(* IEC 61131-3 sources: daoli-st-library/DL_Base (part 19) *)

(* ---- FB_DL_Vote2oo3.st ---- *)
(*==============================================================================
 * 组件名称 (Component)  : FB_DL_Vote2oo3
 * 所属子库 (Sublibrary) : DL_Base
 * 当前版本 (Version)    : 1.0.0
 * 兼容性   (Platform)   : CODESYS 3.5+ / TwinCAT 3 / 汇川 InoProShop / 施耐德 Machine Expert
 *                         仅依赖 Standard.library（TON / R_TRIG / ABS），零厂商私有库
 * 功能描述 (Function)   : 三通道二取二表决（2oo3）。逐拍统计健康通道数 nHealthy 与
 *                         健康通道中为真的个数 nTrue：
 *                         ① nHealthy >= 3 → 三取二多数表决（2/3 即通过）；
 *                         ② nHealthy = 2 → 降级 1oo2，两健康通道一致才通过，不一致判失配；
 *                         ③ nHealthy <= 1 → 健康数不足，输出保守 FALSE 并置故障；
 *                         ④ 失配须连续维持 tMismatchTime（默认 T#300MS）才判故障，
 *                            消除单拍抖动造成的误判（确认窗消除法）。
 *                         输出同意数 nAgreeCount = 多数派票数 = MAX(nTrue, nHealthy - nTrue)。
 * 接口     (Interface)  : 输入 bCh1/bCh2/bCh3 三通道原始值、bHealthy1/bHealthy2/bHealthy3
 *                         通道健康位、tMismatchTime 失配确认时间、tConfirmTime 健康数不足
 *                         确认时间、bReset 复位电平；输出 bOut 表决结果、nAgreeCount 同意数、
 *                         eState 相位、eCause 成因、bError 故障标志、nErrId 事件码。
 * 边界     (Boundary)   : ① 组态闸：tMismatchTime <= T#0S 或 tConfirmTime <= T#0S → 故障锁存；
 *                         ② 安全侧：任何故障相 bOut 强制 FALSE（保守关断侧），nAgreeCount 置 0；
 *                         ③ TON 两枚 + R_TRIG 一枚在段 0 无条件周期刷新，IN 由当拍判据派生；
 *                         ④ 故障相迁出唯一路径 = bReset 上升沿；⑤ 零全局耦合（无 GVL / 无物理地址）。
 * 解除式   (Release)    : bReset 上升沿 ∧ 组态合法 ∧ tonMismatch.Q = FALSE ∧
 *                         tonInsuff.Q = FALSE ∧ nHealthy >= 2（全为当拍量，R240 范式）。
 *                         自证可满足（终审两式 1）：故障相下两枚 TON 的 IN 仍由当拍判据
 *                         派生，三通道恢复一致且健康数恢复 >= 2 时两 Q 必落假，解除式必可达。
 * 码表     (Codes)      : 16#0001_03EA 故障级：表决故障总码（组态非法 / 通道失配 / 健康数不足），
 *                         锁存至 bReset 上升沿，归因由 eCause 独立成员承载（R190 单件单总码）；
 *                         16#0001_04AD 信息级：降级 1oo2 表决中（健康数恰为 2，无故障）。
 *                         加码反证（R90）：降级 1oo2 与「三通道全健康」在 bOut/nAgreeCount 上
 *                         可同值（nHealthy=2 且一致时 nAgreeCount=2），但二者故障处置不同，
 *                         现有输出组合无法唯一还原「当前仅两通道可信」，故立此信息码。
 *                         码段说明：0001 段故障子带 03xx / 信息子带 04xx，本件取 03EA / 04AD
 *                         （源码实扫该两槽为空，续接同子带已用最大值，未回填碎片孔洞）。
 * 开源溯源 (Origin)     : 道莅自研 clean-room（参考 2oo3 表决结构惯例与参数域，零代码行复制）
 * 修订历史 (Revision)   : 2026-11-19  v1.0.0  R45 首版（批次 1 · 序号 1）
 *==============================================================================*)

TYPE E_DL_V23State :
(
    eIdle  := 0,     // 未使能待运行（健康通道数不足前不输出） / Idle, not enough healthy channels
    eRun   := 10,    // 表决运行 / Voting in progress
    eFault := 90     // 故障锁存相 / Fault latched phase
);
END_TYPE

TYPE E_DL_V23Cause :
(
    eNone       := 0,   // 无故障成因 / No cause
    eCfgIllegal := 1,   // 组态非法 / Illegal configuration
    eMismatch   := 2,   // 健康通道表决失配（确认时间到） / Healthy channels mismatch confirmed
    eInsuff     := 3    // 健康通道数不足（<= 1） / Insufficient healthy channels
);
END_TYPE

FUNCTION_BLOCK FB_DL_Vote2oo3
VAR_INPUT
    bCh1          : BOOL := FALSE;            // 通道 1 原始值 [-] / Channel 1 raw value
    bCh2          : BOOL := FALSE;            // 通道 2 原始值 [-] / Channel 2 raw value
    bCh3          : BOOL := FALSE;            // 通道 3 原始值 [-] / Channel 3 raw value
    bHealthy1     : BOOL := TRUE;             // 通道 1 健康位，FALSE 表示该通道不参与表决 [-] / Channel 1 health, FALSE excludes it
    bHealthy2     : BOOL := TRUE;             // 通道 2 健康位，FALSE 表示该通道不参与表决 [-] / Channel 2 health, FALSE excludes it
    bHealthy3     : BOOL := TRUE;             // 通道 3 健康位，FALSE 表示该通道不参与表决 [-] / Channel 3 health, FALSE excludes it
    tMismatchTime : TIME := T#300MS;          // 失配确认时间，域 > T#0S [ms] / Mismatch confirm time, domain > T#0S
    tConfirmTime  : TIME := T#500MS;          // 健康数不足确认时间，域 > T#0S [ms] / Insufficient-health confirm time
    bReset        : BOOL := FALSE;            // 复位命令，上升沿清故障 [-] / Reset command, rising edge clears fault
END_VAR
VAR_OUTPUT
    bOut          : BOOL;                     // 表决结果，故障相强制 FALSE（安全侧） [-] / Voting result, forced FALSE in fault
    nAgreeCount   : INT;                      // 多数派同意票数 [票] / Majority agreement count [votes]
    eState        : E_DL_V23State;            // 状态出口，段 6 单点映射 / State outlet, single mapping point
    eCause        : E_DL_V23Cause;            // 故障成因出口（R190 归因唯一） / Fault cause outlet
    bError        : BOOL;                     // 故障锁存标志 [-] / Fault latch flag
    nErrId        : UDINT;                    // 事件码，0 = 无事件 / Event code, 0 = no event
END_VAR
VAR
    _eState       : E_DL_V23State := E_DL_V23State.eIdle;      // 内部相位（CASE 唯一写入目标） / Internal phase
    _eCause       : E_DL_V23Cause := E_DL_V23Cause.eNone;      // 故障成因锁存（锁存量） / Latched cause
    tonMismatch   : TON;                      // 失配确认计时，段 0 无条件调用 / Mismatch confirm timer
    tonInsuff     : TON;                      // 健康数不足确认计时，段 0 无条件调用 / Insufficient-health timer
    rtReset       : R_TRIG;                   // 复位沿实例，段 0 无条件调用 / Reset edge instance
    _nHealthy     : INT;                      // 健康通道数当拍量 [路] / Healthy channel count this scan
    _nTrue        : INT;                      // 健康通道中为真的个数当拍量 [路] / TRUE count among healthy channels
    _bDisagree    : BOOL;                     // 健康通道失配当拍量 [-] / Healthy channels disagree
    _bInsuff      : BOOL;                     // 健康数不足当拍量 [-] / Insufficient healthy channels
    _bCfgBad      : BOOL;                     // 组态非法当拍量 [-] / Illegal configuration
    _bFault       : BOOL;                     // 故障锁存位（锁存量） / Latched fault bit
    _uFault       : UDINT;                    // 故障码锁存（锁存量） / Latched fault code
    _uInfo        : UDINT;                    // 信息码，每拍重算 / Info code, recomputed each scan
END_VAR

(* —— 段 0：当拍判据派生 + 定时器与沿实例无条件周期刷新 —— *)
_nHealthy := 0;                                                              // 健康计数起点 0 / Healthy count start
_nTrue    := 0;                                                              // 真票计数起点 0 / TRUE vote count start
IF bHealthy1 THEN                                                            // 通道 1 健康则纳入 / Channel 1 counted if healthy
    _nHealthy := _nHealthy + 1;                                              // 健康数累加 / Accumulate healthy count
    IF bCh1 THEN
        _nTrue := _nTrue + 1;                                                // 真票累加 / Accumulate TRUE vote
    END_IF
END_IF
IF bHealthy2 THEN                                                            // 通道 2 健康则纳入 / Channel 2 counted if healthy
    _nHealthy := _nHealthy + 1;
    IF bCh2 THEN
        _nTrue := _nTrue + 1;
    END_IF
END_IF
IF bHealthy3 THEN                                                            // 通道 3 健康则纳入 / Channel 3 counted if healthy
    _nHealthy := _nHealthy + 1;
    IF bCh3 THEN
        _nTrue := _nTrue + 1;
    END_IF
END_IF
_bDisagree := (_nHealthy >= 2) AND (_nTrue > 0) AND (_nTrue < _nHealthy);     // 健康通道内既有真也有假即失配 / Disagreement inside healthy set
_bInsuff   := (_nHealthy <= 1);                                               // 健康数 <= 1 即不足 / Less than two healthy channels
_bCfgBad   := (tMismatchTime <= T#0S) OR (tConfirmTime <= T#0S);              // 组态非法当拍量 / Illegal configuration this scan
rtReset(CLK := bReset);                                                      // 复位沿，每拍必调（R228A） / Reset edge, called every scan
tonMismatch(IN := _bDisagree, PT := tMismatchTime);                          // 失配确认计时 / Mismatch confirm timer
tonInsuff(IN := _bInsuff, PT := tConfirmTime);                               // 健康数不足确认计时 / Insufficient-health timer

(* —— 段 1：单拍量预清零（锁存量与 TON/R_TRIG 实例不入清单，R107） —— *)
_uInfo      := 16#0000_0000;          // 信息码每拍重算 / Info recomputed every scan
bOut        := FALSE;                 // 表决结果缺省 FALSE（安全侧） / Result default FALSE, safe side
nAgreeCount := 0;                     // 同意数缺省 0 / Agreement count default 0
nErrId      := 16#0000_0000;          // 事件码缺省无事件 / Event code default none
bError      := FALSE;                 // 故障标志每拍预清，由故障分支同拍置位（R45 配对） / Flag preset, set by fault branch

(* —— 段 2：复位沿 + 组态域闸 —— *)
IF rtReset.Q THEN                                                    // rtReset.Q 为当拍量 / current-scan edge
    _bFault := FALSE;                                                // 清故障锁存位（锁存量） / Clear fault latch
    _uFault := 16#0000_0000;                                         // 清故障锁存码（锁存量） / Clear latched code
    _eCause := E_DL_V23Cause.eNone;                                  // 清成因（锁存量） / Clear latched cause
    IF _eState = E_DL_V23State.eFault THEN
        _eState := E_DL_V23State.eIdle;                              // 故障相迁出唯一路径 / Sole exit from fault phase
    END_IF
END_IF
IF _bCfgBad THEN                                                     // 组态域闸 / Configuration gate
    _uFault := 16#0001_03EA;                                         // 故障级：表决故障总码 / Fault-level: voting fault code
    _bFault := TRUE;                                                 // 锁存置位 / Latch set
    bError  := TRUE;                                                 // 故障标志同拍置位（R45 配对） / Error flag set same scan
    _eCause := E_DL_V23Cause.eCfgIllegal;                            // 归因：组态非法 / Cause: illegal configuration
END_IF

(* —— 段 3：失配与健康数不足（确认窗到时才判，消除单拍抖动） —— *)
IF (NOT _bFault) AND tonMismatch.Q THEN                              // 失配确认窗到 / Mismatch confirm elapsed
    _uFault := 16#0001_03EA;
    _bFault := TRUE;
    bError  := TRUE;
    _eCause := E_DL_V23Cause.eMismatch;                              // 归因：通道失配 / Cause: channel mismatch
END_IF
IF (NOT _bFault) AND tonInsuff.Q THEN                                // 健康数不足确认窗到 / Insufficient-health elapsed
    _uFault := 16#0001_03EA;
    _bFault := TRUE;
    bError  := TRUE;
    _eCause := E_DL_V23Cause.eInsuff;                                // 归因：健康数不足 / Cause: insufficient health
END_IF

(* —— 段 4：故障解除式（R240 全当拍量） —— *)
IF rtReset.Q AND (NOT _bCfgBad) AND (NOT tonMismatch.Q) AND (NOT tonInsuff.Q) AND (_nHealthy >= 2) THEN
    _bFault := FALSE;                                                // 清故障锁存位（锁存量） / Clear fault latch
    _uFault := 16#0000_0000;                                         // 清故障锁存码（锁存量） / Clear latched code
    _eCause := E_DL_V23Cause.eNone;                                  // 清成因（锁存量） / Clear latched cause
END_IF

(* —— 段 4A：故障锁存相位迁移闸 —— *)
IF _bFault AND (_eState <> E_DL_V23State.eFault) THEN                // 锁存即入故障相 / Latch enters fault phase
    _eState := E_DL_V23State.eFault;
END_IF

(* —— 段 5：相位机（ENUM 全成员显式标签 + ELSE 兜底，R128） —— *)
CASE _eState OF

E_DL_V23State.eIdle:
    IF (_nHealthy >= 2) AND (NOT _bFault) THEN                        // 出口 1：健康通道恢复 / Enough healthy channels
        _eState := E_DL_V23State.eRun;                                // 进表决运行 / Enter voting run
    ELSIF _bFault THEN                                                // 出口 2：已锁故障（前置被破坏） / Fault latched
        _eState := E_DL_V23State.eFault;
    END_IF

E_DL_V23State.eRun:
    IF _nHealthy < 2 THEN                                             // 出口 1：健康数跌破 2 / Healthy count drops below two
        _eState := E_DL_V23State.eIdle;                               // 退回未使能待恢复 / Back to idle awaiting recovery
    ELSIF _bFault THEN                                                // 出口 2：故障锁存 / Fault latched
        _eState := E_DL_V23State.eFault;
    END_IF

E_DL_V23State.eFault:
    ;                                                                 // 故障相：仅段 4 复位沿可迁出 / Only the reset edge leaves this phase

ELSE
    _uFault := 16#0001_03EA;                                          // 故障级：非法相位兜底（归并总码） / Illegal-phase fallback
    _bFault := TRUE;                                                  // 锁存置位 / Latch set
    bError  := TRUE;                                                  // 故障标志同拍置位（R45 配对） / Error flag set same scan
    _eCause := E_DL_V23Cause.eCfgIllegal;                             // 归因：相位非法归并组态 / Cause: phase illegal mapped to config
    _eState := E_DL_V23State.eFault;                                  // 强制回故障相 / Force fault phase

END_CASE

(* —— 段 6：出口单点映射（名实同源；锁存码回放） —— *)
IF _bFault THEN
    bOut        := FALSE;                                             // 故障相保守关断侧 / Conservative OFF in fault
    nAgreeCount := 0;                                                 // 故障相同意数置 0 / Agreement count zeroed in fault
ELSE
    IF (_nTrue * 2) > _nHealthy THEN                                  // 多数派为真（严格过半） / Strict majority TRUE
        bOut := TRUE;
    ELSE
        bOut := FALSE;                                                // 无过半多数（含 1oo2 不一致）保守 FALSE / No majority, conservative FALSE
    END_IF
    IF _nTrue >= (_nHealthy - _nTrue) THEN                            // 多数派票数 = MAX(真, 假) / Majority votes
        nAgreeCount := _nTrue;
    ELSE
        nAgreeCount := _nHealthy - _nTrue;
    END_IF
    IF _nHealthy = 2 THEN                                             // 降级 1oo2 运行（信息级） / Degraded 1oo2 operation
        _uInfo := 16#0001_04AD;
    END_IF
END_IF
IF _bFault THEN
    nErrId := _uFault;                                                // 故障锁存码回放 / Replay latched fault code
ELSE
    nErrId := _uInfo;                                                 // 信息码 / Info code
END_IF
bError := _bFault;                                                    // 故障标志与锁存同源（名实双出口，R191） / Flag from latch
eState := _eState;                                                    // 状态出口 / State outlet
eCause := _eCause;                                                    // 成因出口 / Cause outlet

END_FUNCTION_BLOCK

(* ---- FB_DL_VoteKooN.st ---- *)
(*
  ==================================================================
  组件名 Component  : FB_DL_VoteKooN
  分类   Category   : DL_Base
  复杂度 Complexity  : cx5
  版本   Version    : 1.0.0
  功能   Purpose    : N 中取 K 安全表决器（MooN 架构）。对 N 个通道的触发量
                      与健康位做 KooN 表决：健康通道中触发数 ≥ K 即表决输出
                      置位；支持通道故障掩码注入（强制剔除指定通道）与 K/N
                      可组态；组态越域锁存故障并输出安全侧。与固定 2oo3 的
                      FB_DL_Vote2oo3 分工互引（固定架构 vs 通用 KooN）。
  来源   Source     : self-std（IEC 61508 MooN 架构公开表决语义）
  溯源   Origin     : IEC 61131-3 标准语义的道莅防御性实现；KooN（MooN）表决
                      为 IEC 61508 公开安全架构语义，clean-room 自研实现，未
                      复制任何厂商私有库源码。
  平台   Platform   : 纯 IEC 61131-3（Standard.library: R_TRIG，无私有库）
  分工声明 Split     : 与 DL_Base 存量 FB_DL_Vote2oo3 分工——Vote2oo3 为固定
                      2oo3 单一架构快捷件，本件为通用 KooN（K 与 N 均可组态，
                      通道数 2..8）架构件；两者不互相替代。
  作者   Author     : 道莅代码库 · PLC 编程专家（R58）
  ------------------------------------------------------------------
  边界 Boundary     :
                      一 组态域：nN ∈ [2..8]，nK ∈ [1..nN]；越域锁存 bCfgBad
                         （解除路径 = bReset 上升沿，且组态恢复后不再重锁），
                         锁存期表决出口置安全侧 TRUE（fail-safe 跳闸，R191
                         显式声明为降级安全值 + 置标志）；
                      二 健康位 FALSE 或掩码注入 TRUE 的通道不计入表决基数；
                         掩码通道的触发量不参与任何判定；
                      三 数组按固定界 0..7 遍历，nN 越界的槽位天然不入基数
                         （无动态下标，结构性越界防御）；
                      四 失能（bEnable = FALSE）输出冻结保持末值（R191 冻结
                         保持声明），组态闸与计数仍每拍刷新；
                      五 无全局变量、无外部变量声明、无物理地址寻址。
  修订记录 Revision  :
    2026-11-21  v1.0.0  R58 首版（批 1 · 序号 1）
  ==================================================================
*)

TYPE E_DL_VknCause :
(
    eNone   := 0, // 无成因 / no cause
    eCfgBad := 1  // 组态非法：N 或 K 越域（故障级，与 bError 配对）/ an illegal config, N or K out of the domain
);
END_TYPE

FUNCTION_BLOCK FB_DL_VoteKooN
VAR_INPUT
    abChnTrip : ARRAY[0..7] OF BOOL; // 通道触发量数组，槽位即通道号 [-] / the channel trip array, the slot is the channel number
    abChnOk   : ARRAY[0..7] OF BOOL; // 通道健康位，FALSE = 通道故障剔除 [-] / the channel health bits, false excludes the faulty channel
    abChnMask : ARRAY[0..7] OF BOOL; // 通道故障掩码注入，TRUE = 强制剔除 [-] / the channel mask injection, true forces the exclusion
    nN        : USINT := 3;   // 表决基数 N（参与通道数）[个]，域 2..8 / the voter base N [channel], two through eight
    nK        : USINT := 2;   // 表决门限 K（跳闸所需触发数）[个]，域 1..N / the voter threshold K [channel], one through N
    bEnable   : BOOL := TRUE; // 使能，失能冻结输出末值 [-] / enable, disabling freezes the outputs
    bReset    : BOOL := FALSE; // 复位上升沿清组态故障锁存 [-] / reset rising edge clears the config fault latch
END_VAR
VAR_OUTPUT
    bTrip    : BOOL := FALSE; // 表决出口，TRUE = 健康通道触发数 ≥ K [-] / the vote outlet, true when the healthy trips reach K
    nHealthy : USINT := 0;    // 参与表决的健康通道数 [个] / the healthy channel count participating [channel]
    nTripChn : USINT := 0;    // 健康通道中的触发通道数 [个] / the tripped channel count among the healthy [channel]
    eCause   : E_DL_VknCause := E_DL_VknCause.eNone; // 成因出口，锁存回放 [枚举] / the cause outlet replayed
    bError   : BOOL := FALSE; // 故障锁存标志（组态越域）[-] / the fault latch flag, a config violation
END_VAR
VAR
    rtReset  : R_TRIG; // 复位沿检测，段 0 无条件刷新 / the reset edge, refreshed unconditionally
    _nI      : DINT;   // 通道遍历索引 [槽] / the channel loop index [slot]
    _nBase   : DINT;   // 参与基数（健康且未掩码）[个] / the participating base [channel]
    _nTrip   : DINT;   // 健康通道触发计数 [个] / the trip count among the healthy [channel]
    _nND     : DINT;   // N 的 DINT 工作副本 [个]（规避 USINT 混型比较）/ the DINT working copy of N [channel]
    _nKD     : DINT;   // K 的 DINT 工作副本 [个] / the DINT working copy of K [channel]
    _bCfgL   : BOOL := FALSE; // 组态故障锁存位 [-] / the config fault latch bit
END_VAR

// 段 0｜沿检测无条件周期刷新（禁入分支）/ segment 0, the unconditional refresh
rtReset(CLK := bReset); // 复位沿 / the reset edge

// 段 1｜复位沿作用域：清组态故障锁存（作用域逐项声明）/ segment 1, the reset edge scope
IF rtReset.Q THEN // 复位沿 / the reset edge
    _bCfgL := FALSE; // 作用域一：清组态锁存 / scope one, clear the config latch
    eCause := E_DL_VknCause.eNone; // 作用域一：清成因 / scope one, clear the cause
END_IF

// 段 2｜组态域闸（边界一）：N ∈ [2..8]，K ∈ [1..N] / segment 2, the config gate
_nND := USINT_TO_DINT(nN); // 升宽比较副本 / the widened comparison copy
_nKD := USINT_TO_DINT(nK); // 升宽比较副本 / the widened comparison copy
IF (nN < 2) OR (nN > 8) OR (nK < 1) OR (nK > nN) THEN // 越域判定（双侧直比，无 ABS）/ the domain verdict, both sides direct
    IF NOT _bCfgL THEN // 未锁存才置位（锁存回放 R152）/ latch only while unlatched
        _bCfgL := TRUE; // 置组态故障锁存 / raise the config fault latch
        eCause := E_DL_VknCause.eCfgBad; // 故障级成因（R45 配对 bError）/ the fault cause
    END_IF
END_IF
bError := _bCfgL; // 故障标志与锁存位同源（R191 名实双出口）/ the flag shares the latch

// 段 3｜通道遍历计数（固定界 0..7，槽位越 nN 的不入基数，边界三）/ segment 3, the channel scan with a fixed bound
_nBase := 0; // 基数清零 / clear the base
_nTrip := 0; // 触发计数清零 / clear the trip count
FOR _nI := 0 TO 7 DO // 固定界循环，无死循环风险 / the fixed bound loop
    IF (_nI < _nND) AND abChnOk[_nI] AND (NOT abChnMask[_nI]) THEN // 在 N 域内且健康且未掩码 / inside N, healthy, and unmasked
        _nBase := _nBase + 1; // 基数推进 / advance the base
        IF abChnTrip[_nI] THEN // 通道触发 / the channel tripped
            _nTrip := _nTrip + 1; // 触发计数推进 / advance the trip count
        END_IF
    END_IF
END_FOR
nHealthy := DINT_TO_USINT(_nBase); // 健康数出口 / the healthy count outlet
nTripChn := DINT_TO_USINT(_nTrip); // 触发数出口 / the trip count outlet

// 段 4｜表决与出口（组态锁存期 fail-safe 置 TRUE，边界一）/ segment 4, the vote and the outlets
IF _bCfgL THEN // 组态故障锁存期 / while the config fault latches
    bTrip := TRUE; // 安全侧跳闸（fail-safe，降级安全值 + bError 置位，R191）/ the fail safe trip with the flag raised
END_IF
IF (NOT _bCfgL) AND bEnable THEN // 组态正常且使能才刷新表决出口 / refresh the vote outlet only when the config is fine and enabled
    bTrip := (_nTrip >= _nKD); // 表决判定：健康触发数 ≥ 门限 K / the vote verdict, the trips reach K
END_IF
// 失能且无组态故障时不进入任何刷新分支：bTrip 冻结保持末值（边界四，R191 冻结保持声明）
// with no config fault and disabled, no refresh branch runs, bTrip freezes at the last value
END_FUNCTION_BLOCK

(* ---- FB_DL_WatchdogMonitor.st ---- *)
(*==============================================================================
 * 组件名称 (Component)  : FB_DL_WatchdogMonitor
 * 所属子库 (Sublibrary) : DL_Base
 * 当前版本 (Version)    : 1.0.0
 * 兼容性   (Platform)   : CODESYS 3.5 / TwinCAT 3 / 汇川 InoProShop / Machine Expert
 *                         仅依赖 Standard.library（TON / R_TRIG）+ 本库双层沿检测构件
 * 功能描述 (Function)   : 外部心跳信号看门狗。监控对象是心跳的"跳变间隔"而不是电平：
 *                         连接还在、脚本已死循环的静默失效工况下，电平永远不变，
 *                         只有跳变间隔能暴露问题。超窗即锁定故障输出并保持，需显式复位；
 *                         同时检测跳变过快（接线抖动 / 心跳被写成恒振荡）并告警，
 *                         该频率告警不锁存，间隔恢复正常即自动消除。
 *                         上电即武装：窗口内没有第一个跳变就按时超时——
 *                         心跳信号必须先证明自己活着，这是刻意设计而非缺陷。
 * 开源溯源 (Origin)     : 原创实现。看门狗的"窗口定时器 + 跳变沿复位"模式为工业界通行做法，
 *                         跳变间隔语义与高频告警为本库差异化设计，未复制任何源码。
 * 本文件内含       : TYPE  E_DL_WdtState（配套枚举，归属 DL_Base）
 *                    FB    FB_DL_WatchdogMonitor
 * 依赖     (Depends)    : FB_DL_DualEdgeTrig（首轮 #2，仅取其电平输出）
 *                         Standard.library: TON / R_TRIG
 * 红线自检 (Redline)    : R1 ✓ 禁用全局存储与物理寻址 ｜ R2 ✓ 无地址直写
 *                         R3 ✓ 纯 IEC 61131-3 ｜ R4 ✓ 窗口钳位 + 零窗口合法性判定
 *                         R5 ✓ 全变量中英双语同行注释 ｜ R6 ✓ 三态 ENUM + CASE + ELSE 兜底
 *                         R7 ✓ 三实例主体最前部无条件刷新 ｜ R8 ✓ 上限与常量全常量化
 *
 * 【依赖收窄留档 / Dependency narrowing（R11）】
 *   规格书 B5 要求跳变计数直接复用双层沿检测构件的上升/下降计数输出。
 *   实测该构件当前版本的上升/下降事件输出以"上一周期电平"做资格与运算，
 *   在真实上升沿那一周期上一周期电平必然为 FALSE，导致事件恒不成立、计数恒不增长。
 *   为避免看门狗核心功能被上游缺陷阻塞，本组件只从该构件取"当前电平"（正确且稳定），
 *   跳变判定与计数在本地以电平差分为准，饱和口径与故障码口径与上游保持一致。
 *   上游修复后可改为直接读其事件输出，届时本段留档同步撤销。
 *   （2026-11-14 终审补注：上游缺陷已在 FB_DL_DualEdgeTrig v1.0.1 修复，
 *     其事件输出恢复正确。本组件继续保留本地电平差分口径——两者行为等价，
 *     且本地派生同时服务于 tSinceToggle 与频率判定，独立于上游事件口更稳；
 *     是否收敛为上游事件输出留待 Level 1 统一重构时评估，本版不改行为。）
 *   The dependency's edge outputs are qualified by the previous level, which makes them
 *   permanently FALSE on a genuine edge. This component therefore consumes only its
 *   level output and derives toggles locally, keeping the same saturation policy.
 *   (Final review note: the upstream defect is fixed in v1.0.1; the local derivation is
 *   kept because it is behaviour-equivalent and also feeds the silence measurement.)
 *
 * 修订历史 (Revision)   :
 *   2026-11-14  v1.0.0  首版入库（Phase 1 第二轮 · Level 0 批次 B）
 *   2026-11-14  v1.0.0  含依赖收窄留档（见上）
 *   2026-11-14  v1.0.0  终审补注依赖收窄现状（仅注释同步，逻辑未变，版本不变）
 *============================================================================*)

(*-----------------------------------------------------------------------------
 * 枚举: E_DL_WdtState（归属 DL_Base，与 FB_DL_WatchdogMonitor 同文件）
 * 含义: 看门狗工作状态。数值步长留空位便于后续插态而不破坏已有工程。
 *----------------------------------------------------------------------------*)
TYPE E_DL_WdtState :
(
    eArmed    := 0,    // 监控中：窗口计时进行，等待下一次跳变 / Armed, the window timer runs and waits for the next toggle
    eFault    := 10,   // 心跳超时锁定：仅复位沿可解除 / Timeout latched, only the reset edge releases it
    eDisabled := 20    // 未启用：输出全清，重新使能视同首次武装 / Disabled, re-enabling behaves like a first arming
);
END_TYPE

FUNCTION_BLOCK FB_DL_WatchdogMonitor
VAR_INPUT
    bHeartbeat   : BOOL;                  // 被监控心跳信号（期望周期性跳变）/ Monitored heartbeat, expected to toggle periodically
    tMaxInterval : TIME := T#2S;          // 最大允许跳变间隔 [ms] / Max allowed toggle interval [ms]
    tMinInterval : TIME := T#5MS;         // 最小合法跳变间隔 [ms]，低于视为异常信号 / Min legal interval [ms], below is abnormal
    bEnable      : BOOL := TRUE;          // 使能 / Enable
    bReset       : BOOL;                  // 上升沿：清除故障并重新武装 / Rising edge: clear fault and re-arm
END_VAR
VAR_OUTPUT
    bAlive       : BOOL;     // 心跳健康（未超时且未触发频率异常）/ Heartbeat healthy, no timeout and no rate anomaly
    bTimeout     : BOOL;     // 心跳超时锁存 / Timeout latched
    tSinceToggle : TIME;     // 距上次跳变的时长 [ms] / Time since the last toggle [ms]
    uToggleCount : UDINT;    // 累计跳变次数 [次]（诊断用）/ Accumulated toggles [count], diagnostics
    bError       : BOOL;     // 故障标志，bReset 清除 / Fault flag, cleared by bReset
    uErrorId     : UDINT;    // 故障码，0 = 无故障 / Error code, 0 = no error
END_VAR
VAR
    fbDual       : FB_DL_DualEdgeTrig;    // 依赖构件实例，仅取电平输出 / Dependency instance, level output only
    fbTonWatch   : TON;                   // 看门狗窗口计时器 / Watchdog window timer
    fbTrigReset  : R_TRIG;                // 复位上升沿检测实例 / Reset rising edge detector instance
    eState       : E_DL_WdtState;         // 主状态机 / Main state machine
    tMinLast     : TIME;                  // 上一次相邻跳变间隔 [ms]（诊断留档）/ Last observed toggle interval [ms]
    bLastLevel   : BOOL;                  // 上周期心跳电平，跳变派生用 / Previous heartbeat level for toggle derivation
    bToggle      : BOOL;                  // 本周期检测到跳变 / Toggle detected in this scan
    tMaxEff      : TIME;                  // 钳位后的窗口 [ms] / Clamped window [ms]
    tPrevSince   : TIME;                  // 上周期末的静默时长 [ms]，间隔测量用 / Silence at the end of the last scan [ms]
    tFrozenSince : TIME;                  // 故障瞬间冻结的静默时长 [ms] / Frozen silence at the fault instant [ms]
    bHasToggled  : BOOL;                  // 是否已观测到过至少一次跳变 / At least one toggle has been observed
    bRateBad     : BOOL;                  // 本周期频率异常（不锁存）/ Rate anomaly this scan, not latched
    bWindowBad   : BOOL;                  // 窗口参数非法 / Illegal window parameter
    bCountSat    : BOOL;                  // 跳变计数饱和标志 / Toggle count saturation flag
    bStateBad    : BOOL;                  // 非法状态命中标志 / Illegal state hit flag
    uToggleLocal : UDINT;                 // 本地跳变计数 [次] / Local toggle counter [count]
END_VAR
VAR CONSTANT
    DL_WDT_INTERVAL_MAX : TIME  := T#1H;            // 窗口上限钳位 [ms] / Window clamp [ms]
    DL_WDT_COUNT_MAX    : UDINT := 16#FFFF_FFFE;    // 跳变计数饱和上限 [次] / Toggle count saturation limit
END_VAR

(*------------------------------------------------------------------------------
 * 段 1｜无条件刷新区（红线 R7）：依赖实例与两个标准实例全部位于主体最前部
 *      Unconditional refresh zone: dependency instance and both standard instances
 *      严禁进入任何 IF / CASE 分支，否则窗口计时会被条件化并失去看门狗意义
 *      No instance call may sit inside IF / CASE, otherwise the window loses its meaning
 *-----------------------------------------------------------------------------*)
fbDual(bSignal := bHeartbeat, bEnable := bEnable, bReset := bReset);
fbTrigReset(CLK := bReset);

(*------------------------------------------------------------------------------
 * 段 2｜跳变派生：电平差分，与跳变计数共用同一个判定源，保证口径唯一
 *      Toggle derivation: level difference, the single source of truth for counting
 *-----------------------------------------------------------------------------*)
bToggle := (fbDual.bLevel AND (NOT bLastLevel)) OR ((NOT fbDual.bLevel) AND bLastLevel);

(*------------------------------------------------------------------------------
 * 段 3｜窗口参数校验（边界 B4）：零窗口视为非法但超时立即受理；超上限钳位
 *      Window validation: a zero window is illegal but honoured as an instant timeout
 *      零窗口意味着"监控无意义"，仍按超时受理以保证输出行为可预期
 *      A zero window is meaningless, yet honouring it keeps the output predictable
 *-----------------------------------------------------------------------------*)
bWindowBad := FALSE;

IF tMaxInterval <= T#0S THEN
    tMaxEff    := T#0S;
    bWindowBad := TRUE;
ELSIF tMaxInterval > DL_WDT_INTERVAL_MAX THEN
    tMaxEff    := DL_WDT_INTERVAL_MAX;
    bWindowBad := TRUE;
ELSE
    tMaxEff    := tMaxInterval;
END_IF

(*------------------------------------------------------------------------------
 * 段 4｜窗口计时（边界 B1）：跳变当周期 IN 断开，ET 自然清零重新起算
 *      Window timing: IN drops on the toggle scan, so ET restarts from zero
 *-----------------------------------------------------------------------------*)
fbTonWatch(IN := (eState = eArmed) AND (NOT bToggle) AND bEnable, PT := tMaxEff);

(*------------------------------------------------------------------------------
 * 段 5｜使能 / 复位 / 主状态机（边界 B2/B6/B7/B8/B9）
 *      Enable, reset and the main state machine
 *-----------------------------------------------------------------------------*)
bRateBad  := FALSE;
bStateBad := FALSE;

IF NOT bEnable THEN
    (*--------------------------------------------------------------------------
     * 段 5a｜使能失效（边界 B6）：输出全清、状态回未启用，跳变计数保留作诊断
     *      Disabled: outputs cleared, state parked; the diagnostic count is kept
     *-------------------------------------------------------------------------*)
    eState       := eDisabled;
    bTimeout     := FALSE;
    bAlive       := FALSE;
    tSinceToggle := T#0S;
    tFrozenSince := T#0S;
    tPrevSince   := T#0S;
    bHasToggled  := FALSE;
    bLastLevel   := fbDual.bLevel;
ELSE
    IF fbTrigReset.Q THEN
        (*----------------------------------------------------------------------
         * 段 5b｜复位（边界 B8）：清故障、回武装、窗口重新起算；不清诊断计数
         *      Reset: clear fault, re-arm, restart the window; the counter is kept
         *---------------------------------------------------------------------*)
        eState       := eArmed;
        bTimeout     := FALSE;
        tFrozenSince := T#0S;
        tPrevSince   := T#0S;
        bHasToggled  := FALSE;
        bLastLevel   := fbDual.bLevel;
    ELSE
        (*----------------------------------------------------------------------
         * 段 5c｜主状态机（红线 R6）：ENUM + CASE + ELSE 兜底
         *      Main state machine with the mandatory ELSE fallback
         *---------------------------------------------------------------------*)
        CASE eState OF

            eDisabled:
                (* 重新使能视同首次武装：不等历史，先要求心跳证明自己活着 *)
                (* Re-enabling behaves like a first arming, the heartbeat must prove itself *)
                eState      := eArmed;
                bHasToggled := FALSE;
                tPrevSince  := T#0S;
                bLastLevel  := fbDual.bLevel;

            eArmed:
                IF bToggle THEN
                    (* 跳变计数（饱和停增，不回绕） *)
                    (* Toggle count, saturating instead of wrapping around *)
                    IF uToggleLocal < DL_WDT_COUNT_MAX THEN
                        uToggleLocal := uToggleLocal + UDINT#1;
                    ELSE
                        bCountSat := TRUE;
                    END_IF

                    (*----------------------------------------------------------
                     * 段 5c-1｜频率异常（边界 B3）：相邻跳变间隔小于下限即告警
                     *      Rate anomaly: an interval below the minimum raises the alarm
                     *      首个跳变不参与判定（尚无参照间隔），间隔为 0 亦不判定
                     *      The first toggle and a zero interval are not qualified
                     *---------------------------------------------------------*)
                    IF bHasToggled AND (tPrevSince > T#0S) AND (tPrevSince < tMinInterval) THEN
                        bRateBad := TRUE;
                    END_IF

                    tMinLast    := tPrevSince;
                    bHasToggled := TRUE;
                END_IF

                (*--------------------------------------------------------------
                 * 段 5c-2｜超时锁定（边界 B2）：窗口期满即锁存，仅复位可解
                 *      Timeout latch: the expired window latches until a reset
                 *-------------------------------------------------------------*)
                IF fbTonWatch.Q THEN
                    eState       := eFault;
                    bTimeout     := TRUE;
                    tFrozenSince := fbTonWatch.ET;
                END_IF

            eFault:
                (* 故障锁存：输出保持，窗口不再计时，等待复位沿 *)
                (* Fault latched: outputs hold, the window stops, waiting for reset *)
                bTimeout := TRUE;

            ELSE
                (* 非法状态拦截：转故障并上报，不做隐式恢复 *)
                (* Illegal state interception: go to fault and report, no implicit recovery *)
                eState       := eFault;
                bTimeout     := TRUE;
                bStateBad    := TRUE;
                tFrozenSince := T#0S;

        END_CASE;
    END_IF
END_IF

(*------------------------------------------------------------------------------
 * 段 6｜静默时长输出（边界 B2 配套）：故障态显示冻结值而非 0，便于现场判断超了多久
 *      Silence output: the fault state shows the frozen value instead of zero
 *-----------------------------------------------------------------------------*)
IF eState = eArmed THEN
    tSinceToggle := fbTonWatch.ET;
ELSIF eState = eFault THEN
    tSinceToggle := tFrozenSince;
ELSE
    tSinceToggle := T#0S;
END_IF

(*------------------------------------------------------------------------------
 * 段 7｜健康与故障输出：健康 = 武装中且无频率异常；故障 = 超时锁存
 *      Health and fault outputs: healthy means armed without a rate anomaly
 *-----------------------------------------------------------------------------*)
bAlive       := (eState = eArmed) AND (NOT bRateBad) AND (NOT bWindowBad);
bError       := bTimeout;
uToggleCount := uToggleLocal;

(*------------------------------------------------------------------------------
 * 段 8｜故障码优先级：非法状态 > 超时 > 频率异常 > 计数饱和 > 参数钳位
 *      Error priority: illegal state, timeout, rate anomaly, saturation, clamp
 *-----------------------------------------------------------------------------*)
IF bStateBad THEN
    uErrorId := 16#0001_0005;
ELSIF bTimeout THEN
    uErrorId := 16#0001_000C;
ELSIF bRateBad THEN
    uErrorId := 16#0001_0008;
ELSIF bCountSat THEN
    uErrorId := 16#0001_0007;
ELSIF bWindowBad THEN
    uErrorId := 16#0001_0001;
ELSE
    uErrorId := 16#0000_0000;
END_IF

(*------------------------------------------------------------------------------
 * 段 9｜历史更新必须放在全部判定之后：先取沿再改历史，否则跳变永远检测不到
 *      History update must come last, otherwise toggles are never detected
 *      tPrevSince 记录周期末静默时长，供下一次跳变时计算间隔
 *      tPrevSince stores the end-of-scan silence for the next interval measurement
 *-----------------------------------------------------------------------------*)
bLastLevel := fbDual.bLevel;
tPrevSince := fbTonWatch.ET;
END_FUNCTION_BLOCK

(* ---- FB_DL_WatchdogPulseMon.st ---- *)
(*==============================================================================
 * 组件名称 (Component)  : FB_DL_WatchdogPulseMon
 * 所属子库 (Sublibrary) : DL_Base
 * 当前版本 (Version)    : 1.0.0
 * 兼容性   (Platform)   : CODESYS 3.5+ / TwinCAT 3 / 汇川 InoProShop / 施耐德 Machine Expert
 *                         仅依赖 Standard.library（TON / R_TRIG），零厂商私有库
 * 功能描述 (Function)   : 外部看门狗脉冲超时判死 + 恢复确认窗，双阈值。
 *                         ① 判死阈值 tDeathTimeout：相邻两个脉冲上升沿的间隔超过该值即判死。
 *                            实现上把"判死计时"的 IN 接到 (NOT 脉冲沿单拍标志)，每来一个脉冲沿
 *                            计时器被复位一次，因此计时器量的正是"距上一沿的静默时长"。
 *                         ② 恢复确认窗 tRecoverConfirm：判死后不因单个脉冲就复生，必须连续
 *                            tRecoverConfirm 内持续有脉冲（即判死计时器始终未被 Q 置起）才恢复。
 *                         判死为锁存量（bDead 保持），恢复是显式二段：eRecover 期间维持 bDead
 *                         为真、bAlive 仍为假，只有确认窗走完才同时翻转——杜绝"单个毛刺脉冲
 *                         宣告复活"的假恢复。
 * 接口     (Interface)  : 输入 bPulse 外部看门狗脉冲、tDeathTimeout 判死超时、tRecoverConfirm
 *                         恢复确认窗、bReset 复位；输出 bAlive 存活（未判死且已过确认窗）、
 *                         bDead 判死锁存、bRecovering 恢复确认中、tSilence 当前静默时长、
 *                         eState / eCause / bError。
 * 边界     (Boundary)   : ① 组态闸：tDeathTimeout <= T#0S、tRecoverConfirm < T#0S 或
 *                         tRecoverConfirm > tDeathTimeout（确认窗长于判死窗会让"恢复"永远
 *                         等不到确认）→ 故障锁存并归因 eCfgIllegal。
 *                         ② 双 TON 均在段 0 无条件周期刷新，且 IN 由当拍判据派生（非外部沿清零），
 *                         符合 R228A：tonDeath 与 tonRecover 的 IN 都是当拍表达式的函数。
 *                         ③ 判死锁存位 _bDead 的清除路径唯一 = 恢复确认窗 Q 置起（bReset 上升沿
 *                         亦可强制清，用于检修旁路），两条路径都在段 5 显式写出（R228B 可迁出）。
 *                         ④ 无 TON 跨相复用：两枚计时器分别服务"判死"与"恢复"，PT 语义成对写死，
 *                         不复用同一实例改 PT。
 *                         ⑤ 零全局耦合（无 GVL / 无 VAR_EXTERNAL / 无物理地址）。
 * 分工声明 (Scope)      : 与 `FB_DL_CycleTimeMeasure`（任务周期测量）分工——那件量任务自身节拍，
 *                         本件判**外部**喂狗脉冲是否还活着，二者不可互替（任务节拍正常而外部
 *                         通讯已死是常见工况）。
 * 来源标签 (Source Tag) : T1-7 ◐（开源参考：硬件看门狗脉冲监测与恢复确认参数域，零代码行复制）
 * 解除式   (Release)    : 恢复确认窗 Q 置起（连续 tRecoverConfirm 内有脉冲）∨ bReset 上升沿。
 *                         自证可满足：确认窗 IN = 判死计时器未超时，只要外部真在喂狗，该 IN 持续
 *                         为真，PT 到即置 Q，不依赖任何锁存量或恒假因子。
 * 码表     (Codes)      : 本件不占用任何全局数字码位。出口为 BOOL（bAlive/bDead/bRecovering/
 *                         bError）+ ENUM（eState / eCause），数字码位待主控收口阶段统一派号。
 * 红线自检 (Redline)    : R1 ✓ 零 GVL/VAR_EXTERNAL ｜ R2 ✓ 零 %I/%Q/%M ｜ R3 ✓ 纯 IEC 61131-3
 *                         R4 ✓ 时间域几何闸 + 无浮点比较 ｜ R5 ✓ 声明逐行同行双语注释
 *                         R6 ✓ ENUM+CASE 含 ELSE ｜ R7 ✓ TON/R_TRIG 段 0 无条件刷新
 * 修订历史 (Revision)   : 2026-11-19  v1.0.0  R46 首版（批次 1 · 序号 4）
 *==============================================================================*)

TYPE E_DL_WpmState :
(
    eIdle      := 0,    // 首拍未收到脉冲，等待首沿 / Awaiting the first pulse edge
    eAlive     := 10,   // 脉冲正常相 / Pulses healthy
    eDead      := 20,   // 判死锁存相（保持 bDead） / Dead latched phase
    eRecover   := 30,   // 恢复确认相（维持 bDead，等待确认窗） / Recovery confirmation phase
    eFault     := 90    // 组态故障相（仅复位沿可迁出） / Configuration fault phase
);
END_TYPE

TYPE E_DL_WpmCause :
(
    eNone        := 0,   // 无故障成因 / No cause
    eCfgIllegal  := 1,   // 组态非法（判死窗非正/确认窗越过判死窗） / Illegal configuration
    eTimeout     := 2,   // 静默超判死窗（外部喂狗已停） / Silence exceeded the death timeout
    eRecoverFail := 3,   // 恢复期中再次超时（恢复被推翻） / Timed out again while recovering
    ePhaseBad    := 4    // 非法相位兜底 / Illegal phase fallback
);
END_TYPE

FUNCTION_BLOCK FB_DL_WatchdogPulseMon
VAR_INPUT
    bPulse           : BOOL := FALSE;      // 外部看门狗脉冲（沿有效，电平宽度无关） [-] / External watchdog pulse, edge triggered
    tDeathTimeout    : TIME := T#500MS;    // 判死超时，域 > T#0S（相邻沿最大间隔） [ms] / Death timeout, max gap between edges, domain > T#0S
    tRecoverConfirm  : TIME := T#2S;       // 恢复确认窗，域 >= T#0S 且 <= tDeathTimeout [ms] / Recovery confirm window, 0..death timeout
    bReset           : BOOL := FALSE;      // 复位/检修旁路，上升沿清判死 [-] / Reset or maintenance bypass, rising edge clears death latch
END_VAR
VAR_OUTPUT
    bAlive     : BOOL;              // 存活（未判死且不在恢复确认中） [-] / Alive, not dead and not confirming
    bDead      : BOOL;              // 判死锁存（恢复期仍为真） [-] / Dead latched, still true while confirming
    bRecovering: BOOL;              // 恢复确认中 [-] / Recovery confirmation in progress
    tSilence   : TIME;              // 距上一脉冲沿的静默时长（当拍量） [ms] / Silence since the last pulse edge [ms]
    eState     : E_DL_WpmState;     // 状态出口 [-] / State outlet
    eCause     : E_DL_WpmCause;     // 故障成因出口（R190 归因唯一） [-] / Fault cause outlet
    bError     : BOOL;              // 故障标志（判死或组态非法） [-] / Error flag, dead or illegal configuration
END_VAR
VAR
    _eState    : E_DL_WpmState := E_DL_WpmState.eIdle;    // 内部相位（CASE 唯一写入目标） / Internal phase
    _eCause    : E_DL_WpmCause := E_DL_WpmCause.eNone;    // 故障成因锁存量 / Latched cause
    tonDeath   : TON;               // 判死计时（IN=非脉冲沿），段 0 无条件调用 / Death timer, unconditional call
    tonRecover : TON;               // 恢复确认计时（IN=判死计时未超时），段 0 无条件调用 / Recovery confirm timer, unconditional call
    rtPulse    : R_TRIG;            // 脉冲沿实例，段 0 无条件调用 / Pulse edge instance
    rtReset    : R_TRIG;            // 复位沿实例，段 0 无条件调用 / Reset edge instance
    _bDead     : BOOL;              // 判死锁存位（锁存量） / Latched dead bit
    _bCfgBad   : BOOL;              // 组态非法当拍量 [-] / Illegal configuration this scan
    _bSeenEdge : BOOL;              // 已收到过首个脉冲沿（锁存量） / First edge seen, latched
    _bRecoverFail : BOOL;           // 恢复期再次超时当拍量 [-] / Timed out again during recovery
END_VAR

(* —— 段 0：判据派生 + 三实例无条件周期刷新 —— *)
_bCfgBad := (tDeathTimeout <= T#0S)                         // 判死窗须为正 / Death window must be positive
         OR (tRecoverConfirm < T#0S)                        // 确认窗不得为负 / Confirm window must not be negative
         OR (tRecoverConfirm > tDeathTimeout);              // 确认窗不得越过判死窗（否则永不恢复） / Confirm window must not exceed death window
rtPulse(CLK := bPulse);                                     // 脉冲沿，每拍必调（R228A） / Pulse edge, called every scan
rtReset(CLK := bReset);                                     // 复位沿，每拍必调 / Reset edge, called every scan
tonDeath(IN := NOT rtPulse.Q, PT := tDeathTimeout);         // 判死计时：每来一个沿即复位（IN 由当拍判据派生，非外部清零） / Death timer reset by each edge
tonRecover(IN := (NOT tonDeath.Q) AND (NOT _bCfgBad), PT := tRecoverConfirm);   // 恢复确认：判死计时未超时即视为在喂狗 / Recovery confirm while pulses keep coming

(* —— 段 1：单拍量预清零（锁存量 _bDead / _bSeenEdge / _eCause 不入清单，R107） —— *)
bAlive      := FALSE;           // 存活位每拍预清 / Alive preset
bDead       := FALSE;           // 判死出口每拍预清，锁存分支同拍回填 / Dead outlet preset
bRecovering := FALSE;           // 恢复位每拍预清 / Recovering preset
bError      := FALSE;           // 故障标志每拍预清（R45 配对） / Error flag preset
tSilence    := T#0S;            // 静默时长每拍预清 / Silence preset

(* —— 段 2：静默时长出口（判死计时器已量出的时长直接回放，不另起计时器） —— *)
IF tonDeath.Q THEN
    tSilence := tDeathTimeout;                  // 已超时：报判死窗值（真实静默 >= 该值，取保守下界） / Timed out: report the death window as a conservative bound
ELSE
    tSilence := T#0S;                           // 未超时：本件不暴露亚阈值静默时长（TON 无 ET 出口依赖，保持跨平台） / Below threshold: not exposed
END_IF

(* —— 段 3：复位沿 / 组态闸 —— *)
IF rtReset.Q THEN
    _bDead := FALSE;                            // 清判死锁存（检修旁路） / Clear dead latch
    _bRecoverFail := FALSE;                     // 清恢复失败标记 / Clear recovery-fail flag
    IF _eState = E_DL_WpmState.eFault THEN
        _eState := E_DL_WpmState.eIdle;         // 故障相迁出（R228B） / Leave fault phase
    END_IF
    IF _eState = E_DL_WpmState.eDead THEN
        _eState := E_DL_WpmState.eIdle;         // 判死相迁出（R228B，第二条可迁出路径） / Leave dead phase, second exit path
    END_IF
END_IF
IF _bCfgBad THEN
    _eState := E_DL_WpmState.eFault;            // 组态非法入故障相 / Illegal configuration enters fault phase
    _eCause := E_DL_WpmCause.eCfgIllegal;       // 归因：组态非法 / Cause: illegal configuration
END_IF

(* —— 段 4：首沿捕获（未见过沿前不判死，避免上电即报死） —— *)
IF rtPulse.Q THEN
    _bSeenEdge := TRUE;                         // 首沿锁存（锁存量） / First edge latched
    IF (_eState = E_DL_WpmState.eIdle) THEN
        _eState := E_DL_WpmState.eAlive;        // 首沿即入存活相 / First edge enters alive phase
    END_IF
END_IF

(* —— 段 5：判死与恢复（判死锁存，恢复二段确认；两条清除路径显式列出） —— *)
_bRecoverFail := (_eState = E_DL_WpmState.eRecover) AND tonDeath.Q;     // 恢复期中再次超时 / Timed out again while recovering
IF (_eState <> E_DL_WpmState.eFault) AND _bSeenEdge AND tonDeath.Q THEN
    _bDead := TRUE;                             // 判死锁存（锁存量） / Latch dead
    _eCause := E_DL_WpmCause.eTimeout;          // 归因：静默超时 / Cause: silence timeout
    IF _eState = E_DL_WpmState.eRecover THEN
        _eCause := E_DL_WpmCause.eRecoverFail;  // 归因：恢复被推翻 / Cause: recovery overturned
        _eState := E_DL_WpmState.eDead;         // 回到判死相 / Back to dead phase
    ELSIF _eState <> E_DL_WpmState.eDead THEN
        _eState := E_DL_WpmState.eDead;         // 首次判死 / First death detection
    END_IF
END_IF
IF _eState = E_DL_WpmState.eDead THEN
    IF tonRecover.Q THEN
        _bDead := FALSE;                        // 清除路径 1：恢复确认窗走完 / Exit path 1: recovery window completed
        _eCause := E_DL_WpmCause.eNone;         // 清成因 / Clear cause
        _eState := E_DL_WpmState.eAlive;        // 回存活相 / Back to alive phase
    ELSIF NOT tonDeath.Q THEN
        _eState := E_DL_WpmState.eRecover;      // 转入恢复确认相（bDead 仍为真） / Enter recovery phase, dead still true
    END_IF
END_IF

(* —— 段 6：相位机（ENUM 全成员显式标签 + ELSE 兜底，R128） —— *)
CASE _eState OF

E_DL_WpmState.eIdle:
    IF _bCfgBad THEN                                        // 出口 1：组态非法 / Illegal configuration
        _eState := E_DL_WpmState.eFault;
    ELSIF _bSeenEdge THEN                                   // 出口 2：已见首沿 / First edge seen
        _eState := E_DL_WpmState.eAlive;
    END_IF

E_DL_WpmState.eAlive:
    IF _bCfgBad THEN                                        // 出口 1：组态转非法 / Configuration went illegal
        _eState := E_DL_WpmState.eFault;
    ELSIF _bDead THEN                                       // 出口 2：判死锁存 / Dead latched
        _eState := E_DL_WpmState.eDead;
    END_IF

E_DL_WpmState.eDead:
    IF _bDead = FALSE THEN                                  // 出口：锁存已清（段 5 两条路径之一） / Latch cleared by one of the two paths
        _eState := E_DL_WpmState.eAlive;
    END_IF

E_DL_WpmState.eRecover:
    IF _bDead = FALSE THEN                                  // 出口：确认窗走完，恢复成立 / Recovery window completed
        _eState := E_DL_WpmState.eAlive;
    ELSIF tonDeath.Q THEN                                   // 出口：恢复被推翻（段 5 已置 _bRecoverFail） / Recovery overturned
        _eState := E_DL_WpmState.eDead;
    END_IF

E_DL_WpmState.eFault:
    ;                                                       // 故障相：仅段 3 复位沿可迁出 / Only the reset edge leaves this phase

ELSE
    _eCause := E_DL_WpmCause.ePhaseBad;                     // 归因：非法相位 / Cause: illegal phase
    _eState := E_DL_WpmState.eFault;                        // 强拉故障相 / Force fault phase

END_CASE

(* —— 段 7：出口单点映射（名实双出口，R191） —— *)
IF _eState = E_DL_WpmState.eFault THEN
    bDead := _bDead;                                        // 故障相回放锁存值（不臆造） / Replay latch in fault phase
ELSE
    bDead := _bDead;                                        // 非故障相同样回放锁存值 / Replay latch outside fault phase
END_IF
bRecovering := (_eState = E_DL_WpmState.eRecover);          // 恢复确认中 / Recovery confirmation in progress
bAlive      := (_eState = E_DL_WpmState.eAlive) AND (NOT _bDead);          // 存活 = 存活相且未锁存 / Alive = alive phase and not latched
bError      := _bDead OR (_eState = E_DL_WpmState.eFault);  // 故障标志 = 判死或组态故障 / Error = dead or configuration fault
eState      := _eState;                                     // 状态出口 / State outlet
eCause      := _eCause;                                     // 成因出口 / Cause outlet

END_FUNCTION_BLOCK

(* ---- FB_DL_BidirectionalCounter.st ---- *)
(*==============================================================================
 * 组件名称 (Component)  : FB_DL_BidirectionalCounter
 * 所属子库 (Sublibrary) : DL_Base
 * 当前版本 (Version)    : 1.0.0
 * 组件分类 (Category)   : 功能块（FUNCTION_BLOCK）· 双向预设计数器 · CTUD 超集
 * 兼容性   (Platform)   : CODESYS 3.5 / TwinCAT 3 / 汇川 InoProShop / Schneider
 *                         Machine Expert；仅依赖 Standard.library 的 R_TRIG
 * 功能描述 (Function)   : 上 / 下双向计数（CU / CD 双沿入口），带装载（Load）、
 *                         复位（Reset）、上下独立预设（PV_UP / PV_DN）与双向
 *                         到预设输出（QU / QD），支持饱和不回绕与同拍双边沿
 *                         「加优先」仲裁。对应 IEC 61131-3 标准 CTUD 语义的
 *                         超集（标准 CTUD 只有单一 PV，本件上下各一个预设）。
 *                         典型场景：库位进出双向计数、双向行程脉冲累计、
 *                         双向流量累积、批次进出料差额核算。
 * 职责矩阵 (Scope map)  : 本库计数四件套职责互斥，不可互相替代：
 *                         FB_DL_EventCounter      通用事件累加（单向、无预设）
 *                         FB_DL_ModuloCounter     取模回绕工位索引（单向、循环）
 *                         FB_DL_PresetCounterSat  单向上下限双预设饱和
 *                         本件                    双向 CU 加 CD，双向独立预设，
 *                                                 双向饱和，加优先仲裁
 * 设计要点 (Key notes)  : ① 执行次序写死：预清零 → 取沿 → 预设校验 → 复位 →
 *                           装载 → 计数 → 饱和 → 比较输出，次序颠倒会出现
 *                           「装载拍还多计一个」这类现场最难查的缺陷；
 *                         ② 装载优先于计数：装载边沿拍内计数分支被完全跳过，
 *                           保证「装载值」不会被同拍计数污染；
 *                         ③ 同拍双边沿按「加优先」处理（净加 1），与 IEC
 *                           CTUD 惯例一致，已在注释中写死，不做方向仲裁参数；
 *                         ④ 预设倒置（PV_UP 小于等于 PV_DN）只锁故障不冻结
 *                           计数，与 FB_DL_PresetCounterSat 的「倒置即冻结」
 *                           策略相反，差异在此显式声明（现场止损优先）；
 *                         ⑤ QU / QD 为保持型（R27）：每拍按当前 CV 重算，
 *                           不允许只在「跨越预设那一拍」置位，否则 HMI 会
 *                           看到输出闪断。
 * 开源溯源 (Origin)     : lgf-counter。参考 LGF（Libre Graphical Framework）
 *                         公开函数库「Counter」分类中双向计数类函数的功能
 *                         分类与参数域（CU / CD / LOAD / PV 四组入口形态），
 *                         只借分类、参数域与命名习惯，算法与实现 100% 自有
 *                         clean-room，不构成衍生作品。
 * 依赖     (Depends)    : 无 DL_ 内部依赖；仅 Standard.library 的 R_TRIG
 * 故障码表 (Error codes):
 *   16#0001_0118【信息级】装载值越界被钳位，装载照常完成
 *   16#0001_0215【故障级】预设倒置（PV_UP 小于等于 PV_DN），锁存 bError，
 *                        计数不冻结；只能由 bReset 清除
 *   16#0001_0216【故障级】保留位，本块无 CASE 主状态机，仅作防御式默认码
 *   信息级码只进 uErrorId，不置 bError（R21）。
 * 验收向量 (Acceptance) :
 *   V1 基本双向：PV_UP = 3 / PV_DN = 0，CU 三拍 → CV = 3、QU = TRUE；
 *      CD 一拍 → CV = 2、QU = FALSE、QD = FALSE
 *   V2 同拍双边沿：CU 与 CD 同拍上升 → CV 净加 1，UP 脉冲为 TRUE，DN 为 FALSE
 *   V3 装载优先：bLoad 与 bCountUp 同拍 → CV 等于装载值，装载脉冲为 TRUE，
 *      加计数脉冲为 FALSE
 *   V4 倒置预设：PV_UP = 5 / PV_DN = 10 → bError = TRUE、码 0215，计数继续
 *   V5 饱和：装载 DL_COUNT_MAX 后 CU 一拍 → CV 不变、AtMax = TRUE、无脉冲
 *   V6 保持语义：QU 为 TRUE 后再 CU 两拍，QU 每拍仍为 TRUE（不得回落）
 * 现场提示 (Field notes):
 *   1 bCountUp / bCountDown 取的是上升沿，编码器 A 相脉冲可直接接入，但
 *     高频脉冲（高于任务频率一半）会丢沿，需先由硬件高速计数模块预处理；
 *   2 bReset 为电平有效且优先级高于装载，复位拍不产生装载脉冲，联锁复位
 *     与装载同时给时以复位为准；
 *   3 bEnable 为 FALSE 时冻结计数并清 QU / QD，但 CV 保持，便于检修时保留
 *     当前值；重新使能后从冻结值继续，不做归零；
 *   4 本块不含回绕行为，计到上限即饱和并置 bAtMax，需要回绕请用
 *     FB_DL_ModuloCounter，不要把两个语义混在一个块里。
 * 红线自检 (Redline)    : R1 零全局变量表与外部变量引用 ｜ R2 零物理地址直写
 *                         R3 纯 IEC 61131-3 ｜ R4 DINT 饱和钳位防溢出
 *                         R5 全变量中英双语同行注释 ｜ R6 无 CASE 主状态机（计数型），
 *                         防御式默认码 0216 保留 ｜ R7 三个 R_TRIG 均在分支外刷新
 * 修订历史 (Revision)   :
 *   2026-11-15  v1.0.0  首版入库（Round 10 · Level 0 计数族回补）
 *============================================================================*)

(*==============================================================================
 * 执行次序总表 (Execution order，写死，不得调整)：
 *   序号 步骤            依赖条件              违反后的典型现场现象
 *   1    单拍脉冲预清零  无                    脉冲跨拍泄漏，上一层多计一次
 *   2    三个沿检测刷新  无                    边沿丢失，计数少一拍
 *   3    首扫初始化      仅首扫一次            初值不确定，首件计数错
 *   4    预设域校验      每拍                  预设改错后无提示，输出恒真
 *   5    复位            电平                  复位不生效或复位拍仍计数
 *   6    装载            装载边沿              装载值被同拍计数污染
 *   7    方向仲裁与计数  使能且非复位非装载    上下同拍时净变化不为 1
 *   8    饱和标志        每拍                  到限位后继续累加，溢出回绕
 *   9    比较输出        每拍                  输出只在跨阈拍有效，HMI 闪断
 *   10   对外镜像        每拍                  输出与内部值不同步
 *============================================================================*)

(*==============================================================================
 * 逐拍推演 (Cycle-by-cycle trace)：
 *   场景 A 基本双向（PV_UP=3，PV_DN=0，CV 初值 0）
 *     拍 1 加计数沿 → 方向仲裁走加分支，CV 由 0 变 1，加脉冲为真，QU 假
 *     拍 2 加计数沿 → CV 由 1 变 2，加脉冲为真，QU 假
 *     拍 3 加计数沿 → CV 由 2 变 3，加脉冲为真，QU 真（3 大于等于 3）
 *     拍 4 无沿     → 输出全部保持，QU 仍真（保持语义，不得回落）
 *     拍 5 减计数沿 → CV 由 3 变 2，减脉冲为真，QU 变假
 *   场景 B 同拍双边沿（PV_UP=100）
 *     拍 1 两路同时上升 → 加优先分支，CV 净加 1，加脉冲真、减脉冲假
 *   场景 C 装载与计数同拍
 *     拍 1 装载沿加计数沿 → 装载先执行，CV 等于装载值，装载脉冲真，
 *          本拍跳过计数分支，加脉冲保持假
 *   场景 D 倒置预设（PV_UP=5，PV_DN=10）
 *     拍 1 校验成立 → 锁故障、码 0215，但计数分支照常执行
 *     拍 2 加计数沿 → CV 由 0 变 1（计数未被冻结）
 *   场景 E 饱和（装载 DL_COUNT_MAX 后加计数一拍）
 *     拍 1 装载 → CV 等于上限
 *     拍 2 加计数沿 → 判 CV 不小于上限，不加、不置脉冲，AtMax 为真
 *============================================================================*)

(*==============================================================================
 * 调用示例 (Instance guide)：
 *   VAR fbSlotCnt : FB_DL_BidirectionalCounter; END_VAR
 *   fbSlotCnt(
 *       bCountUp   := bPartInPulse,      // 进料光电脉冲
 *       bCountDown := bPartOutPulse,     // 出料光电脉冲
 *       bLoad      := bRecipeLoad,       // 配方切换时装载
 *       nLoadValue := nRecipeStartCount, // 配方起始值
 *       bReset     := bShiftReset,       // 班次复位
 *       nPresetUp  := nFullLevel,        // 满仓阈值
 *       nPresetDn  := nEmptyLevel,       // 空仓阈值
 *       bEnable    := bStationEnabled);
 *   bFull  := fbSlotCnt.bQu;
 *   bEmpty := fbSlotCnt.bQd;
 *   IF fbSlotCnt.bError THEN nAlarm := fbSlotCnt.uErrorId; END_IF
 *   注意：本块每拍必须调用一次，跳过调用会使边沿检测失效并冻结计数。
 *============================================================================*)

(*==============================================================================
 * 与标准 CTUD 的差异声明 (Deviation from IEC CTUD)：
 *   1 标准 CTUD 只有单一 PV 与单一 QU；本件有上下两个独立预设与两个输出，
 *     以满足双向工艺（满仓与空仓两个阈值）的实际需要；
 *   2 标准 CTUD 在到达计数类型边界时行为未定义；本件在远离边界的
 *     正负二十一万万处饱和，保证加一与减一永不溢出；
 *   3 标准 CTUD 不定义同拍双边沿的净效果；本件写死为加优先净加一；
 *   4 标准 CTUD 无故障概念；本件在预设倒置时锁故障但不冻结计数。
 *============================================================================*)

(*==============================================================================
 * 输出真值表 (Output truth table)：
 *   状态组合                                      QU    QD    含义
 *   使能 且 CV 大于等于 PV_UP                     真    按 QD 判定   满仓侧到达
 *   使能 且 CV 小于等于 PV_DN                     按 QU   真         空仓侧到达
 *   使能 且 PV_UP 大于 CV 大于 PV_DN              假    假         正常区间
 *   失能 且 CV 任意                               假    假         冻结，CV 保持
 *   复位拍 且 CV 归零                             按新 CV 重算        复位优先
 *   PV_UP 与 PV_DN 倒置                           仍按比较式输出      计数不冻结，另报故障
 *   注：两行「按 QU 判定」表示该列的取值与另一列同时成立时互不影响，
 *       两个输出互相独立，不互斥，也不做优先级仲裁。
 *============================================================================*)

(*==============================================================================
 * 参数域与默认值说明 (Parameter domain)：
 *   bCountUp    布尔，上升沿有效；无默认，必须由现场光电或编码器给出
 *   bCountDown  布尔，上升沿有效；无默认，必须由现场光电或编码器给出
 *   bLoad       布尔，上升沿有效；建议用配方切换脉冲或手动装载按钮
 *   nLoadValue  双整数，默认 0，域正负二十一万万；越界自动钳位并置 0118
 *   bReset      布尔，电平有效；建议接班次复位或工位初始化，不接急停
 *   nPresetUp   双整数，默认 100，域建议放在工艺允许范围内，须大于 PV_DN
 *   nPresetDn   双整数，默认 0，域建议放在工艺允许范围内，须小于 PV_UP
 *   bEnable     布尔，默认真；检修时置假可冻结计数并保留当前值
 *   说明：预设值不做内部钳位，只做倒置校验，因为预设是工艺参数而不是
 *   物理量，钳位会掩盖组态错误；倒置只锁故障不改值，便于工程师看到原始填错
 *   的两个数字再决定怎么改。
 *============================================================================*)

(*==============================================================================
 * 常见误用与现场提示 (Field notes)：
 *   1 把高频编码器脉冲直接接到 bCountUp：本块按任务周期取沿，脉冲频率
 *     高于任务频率一半时会丢沿，表现为「计数偏小且不稳定」；正确做法是
 *     先用硬件高速计数模块预处理，或把本块放在高速任务里；
 *   2 把 bReset 接急停回路：急停应当切断输出侧并由安全层处理，本块的复位
 *     只是计数归零，接急停会导致「拍下急停后计数清零」这种不可追溯的行为；
 *   3 把 QU 与 QD 当作互斥的两个状态：两者可能同时为真（当预设区间被
 *     配置成重叠甚至倒置时），上位必须按「两个独立阈值」处理；
 *   4 用本块做取模回绕（如工位号循环）：本块饱和不回绕，请改用
 *     FB_DL_ModuloCounter，两者语义不同，混用会出现「到顶后卡住」；
 *   5 装载后立刻读 CV：装载在同一扫描周期已经完成，读到的就是装载值，
 *     不需要等下一拍；装载脉冲只在该拍为真，下一拍自动清零。
 *============================================================================*)

(*==============================================================================
 * 选型指引 (Which counter to use)：
 *   现场需求                                     应当选用的组件
 *   只想知道「发生了多少次」，不设阈值            FB_DL_EventCounter
 *   工位号在固定范围内循环（如转盘十六工位）      FB_DL_ModuloCounter
 *   单向计数，上下两个阈值，到顶后冻结            FB_DL_PresetCounterSat
 *   双向计数（进出两个方向），上下两个独立阈值    本件
 *   需要计长、累计流量、累计运行时间的工程量      不属于计数件，请用相应工艺件
 *   选错件的典型后果：用本件做转盘循环会在到顶后卡住；用取模件做满仓判断
 *   会永远等不到「满」这个状态，因为取模件根本不产生阈值输出。
 *============================================================================*)

(*==============================================================================
 * 联调清单 (Commissioning checklist)：
 *   1 先确认两路计数信号在静止时都为假，若有常真信号，上电首拍就会误计一次；
 *   2 手动触发一次进料，观察 bUpPulse 是否只闪一拍，若连续闪多拍说明输入
 *     信号抖动，请在上一层加防抖（FC_DL_SignalDebounce 或 FB_DL_SignalDebounce）；
 *   3 把 PV_UP 临时设成当前值，确认 QU 立刻变真，验证比较链路通畅；
 *   4 把 PV_DN 设成大于 PV_UP 的值，确认 bError 置位且码为 0215，验证倒置
 *     保护；验证完毕后必须改回正确值并给一次复位，否则故障锁存不会自清；
 *   5 装载一次上限值再手动加计数，确认 CV 不动且 AtMax 为真，验证饱和；
 *   6 断使能一拍，确认 CV 保持且 QU 与 QD 都为假，验证冻结语义。
 *============================================================================*)

(*==============================================================================
 * 执行代价 (Cost)：
 *   每拍固定两次边沿检测、最多两次整数加减、四次比较，无条件分支以外的
 *   逻辑量恒定，最坏执行时间可静态界定。本件不含循环、不含定时器、不含
 *   浮点，因此放在高速计数中断所挂的任务里也不会有抖动；唯一的库依赖是
 *   R_TRIG，其内部只保存一个上一拍电平，无任何时间量参与。
 *============================================================================*)

FUNCTION_BLOCK FB_DL_BidirectionalCounter
VAR_INPUT
    bCountUp   : BOOL;               // 加计数输入，上升沿加 1，主周期无条件取沿 [-] / Count-up input, rising edge increments by one
    bCountDown : BOOL;               // 减计数输入，上升沿减 1，与加计数同拍时加优先 [-] / Count-down input, rising edge decrements by one
    bLoad      : BOOL;               // 装载请求，上升沿装载，装载拍跳过计数 [-] / Load request, rising edge loads and skips counting
    nLoadValue : DINT := 0;          // 装载值，域 DL_COUNT_MIN 到 DL_COUNT_MAX [计数值] / Load value, range DL_COUNT_MIN to DL_COUNT_MAX
    bReset     : BOOL;               // 复位请求，电平有效：CV 归 0、清 QU / QD 与锁存 [-] / Reset request, level active: CV to zero, clears flags and latches
    nPresetUp  : DINT := 100;        // 加预设值 PV_UP，CV 大于等于此值时 QU 为 TRUE [计数值] / Preset up, QU is TRUE while CV is greater or equal
    nPresetDn  : DINT := 0;          // 减预设值 PV_DN，CV 小于等于此值时 QD 为 TRUE [计数值] / Preset down, QD is TRUE while CV is less or equal
    bEnable    : BOOL := TRUE;       // 使能，FALSE 时冻结计数并清 QU / QD，CV 保持 [-] / Enable, FALSE freezes counting and clears QU and QD
END_VAR
VAR_OUTPUT
    nCv        : DINT;               // 当前计数值 CV，饱和域内不回绕 [计数值] / Current count value, saturated, no wrap-around
    bQu        : BOOL;               // 加预设到达，保持型，CV 大于等于 PV_UP 期间持续为真 [-] / Up preset reached, holding type
    bQd        : BOOL;               // 减预设到达，保持型，CV 小于等于 PV_DN 期间持续为真 [-] / Down preset reached, holding type
    bAtMax     : BOOL;               // 已达上限饱和，再加 1 被拒 [-] / Upper saturation reached, further increments rejected
    bAtMin     : BOOL;               // 已达下限饱和，再减 1 被拒 [-] / Lower saturation reached, further decrements rejected
    bUpPulse   : BOOL;               // 本次实际加计数成功，单拍脉冲 [-] / Increment actually applied this cycle, single-cycle pulse
    bDnPulse   : BOOL;               // 本次实际减计数成功，单拍脉冲 [-] / Decrement actually applied this cycle, single-cycle pulse
    bLoadDone  : BOOL;               // 装载完成，单拍脉冲 [-] / Load completed, single-cycle pulse
    uErrorId   : UDINT;              // 事件码，0 = 无事件 / Event code, 0 = no event
    bError     : BOOL;               // 故障锁存，仅故障级码置位，复位清除 [-] / Fault latch, set only by fault-level codes
END_VAR
VAR
    fbTrigUp    : R_TRIG;            // 加计数边沿检测实例，分支外无条件刷新 [-] / Rising edge detector for count-up input
    fbTrigDown  : R_TRIG;            // 减计数边沿检测实例，分支外无条件刷新 [-] / Rising edge detector for count-down input
    fbTrigLoad  : R_TRIG;            // 装载边沿检测实例，分支外无条件刷新 [-] / Rising edge detector for load request
    bInit       : BOOL := FALSE;     // 首扫标志，初值 FALSE，判据 NOT bInit（R19 范式）[-] / First-scan flag, initial FALSE, tested with NOT
    nCvInt      : DINT := 0;         // 内部计数值，对外经 nCv 镜像输出 [计数值] / Internal count value, mirrored to nCv
    bPresetBad  : BOOL;              // 预设倒置锁存，PV_UP 小于等于 PV_DN 时为 TRUE [-] / Preset inversion latch
    nLoadClamp  : DINT;              // 装载值钳位中间量 [计数值] / Clamped load value temp
END_VAR
VAR CONSTANT
    DL_COUNT_MAX : DINT := 2147483000;   // 计数上限，留安全裕度防加 1 溢出 [计数值] / Count upper bound with overflow margin
    DL_COUNT_MIN : DINT := -2147483000;  // 计数下限，留安全裕度防减 1 溢出 [计数值] / Count lower bound with underflow margin
END_VAR

(*------------------------------------------------------------------------------
 * 段 1｜单拍输出预清零（R25 律①）：三个脉冲输出必须在主体最前部清零
 *      Single-cycle output pre-clear (R25 rule 1): clear the three pulses first
 *      若把清零放在计数之后，上一拍的脉冲会残留到本拍，形成「跨拍泄漏」
 *-----------------------------------------------------------------------------*)
bUpPulse  := FALSE;
bDnPulse  := FALSE;
bLoadDone := FALSE;

(*------------------------------------------------------------------------------
 * 段 2｜边沿实例无条件周期刷新（R7 红线）：不得放在 IF 或 CASE 分支内
 *      Edge instances refreshed unconditionally every cycle, never inside a branch
 *-----------------------------------------------------------------------------*)
fbTrigUp(CLK := bCountUp);
fbTrigDown(CLK := bCountDown);
fbTrigLoad(CLK := bLoad);

(*------------------------------------------------------------------------------
 * 段 3｜首扫初始化（R19 唯一合法范式）：初值 FALSE，判据 NOT bInit
 *      First-scan initialisation: initial value FALSE, tested with NOT bInit
 *      首扫只装载初值与清锁存，不做任何输入相关的动作
 *-----------------------------------------------------------------------------*)
IF NOT bInit THEN
    nCvInt     := 0;                 // 计数从 0 起
    bPresetBad := FALSE;             // 清预设倒置锁存
    bError     := FALSE;             // 清故障锁存
    uErrorId   := 16#0000_0000;      // 清事件码
    bAtMax     := FALSE;             // 饱和位复位
    bAtMin     := FALSE;             // 饱和位复位
    bInit      := TRUE;              // 首扫只做一次
END_IF

(*------------------------------------------------------------------------------
 * 段 4｜预设域校验（每拍重算）：倒置即锁故障，但计数继续
 *      Preset domain check every cycle: inversion latches a fault, counting goes on
 *      现场取舍：宁可带着一组错预设继续计数，也不因一次组态失误停线；
 *      与 FB_DL_PresetCounterSat 的「倒置冻结」策略相反，此处显式声明差异
 *-----------------------------------------------------------------------------*)
IF nPresetUp <= nPresetDn THEN
    bPresetBad := TRUE;
    bError     := TRUE;              // 故障级：锁存
    uErrorId   := 16#0001_0215;
END_IF

(*------------------------------------------------------------------------------
 * 段 5｜复位（电平有效，优先于装载）：CV 归 0，清全部锁存
 *      Reset is level active and takes precedence over load
 *-----------------------------------------------------------------------------*)
IF bReset THEN
    nCvInt     := 0;
    bPresetBad := FALSE;
    bError     := FALSE;
    uErrorId   := 16#0000_0000;
END_IF

(*------------------------------------------------------------------------------
 * 段 6｜装载（边沿有效，优先于计数）：装载拍完全跳过计数分支
 *      Load on rising edge, takes precedence over counting for that cycle
 *      装载值先钳位再落盘，越界只置信息级码，装载动作照常完成
 *-----------------------------------------------------------------------------*)
IF fbTrigLoad.Q AND (NOT bReset) THEN
    nLoadClamp := nLoadValue;
    IF nLoadClamp > DL_COUNT_MAX THEN
        nLoadClamp := DL_COUNT_MAX;
        uErrorId   := 16#0001_0118;  // 装载值越界钳位（信息级）
    ELSIF nLoadClamp < DL_COUNT_MIN THEN
        nLoadClamp := DL_COUNT_MIN;
        uErrorId   := 16#0001_0118;  // 装载值越界钳位（信息级）
    END_IF
    nCvInt    := nLoadClamp;
    bLoadDone := TRUE;               // 装载脉冲，单拍
END_IF

(*------------------------------------------------------------------------------
 * 段 7｜方向仲裁与计数（装载拍与复位拍均不计数）
 *      Direction arbitration and counting, skipped on load and reset cycles
 *      同拍双边沿：加优先，净加 1（IEC CTUD 惯例，语义写死不再开放参数）
 *-----------------------------------------------------------------------------*)
IF bEnable AND (NOT bReset) AND (NOT fbTrigLoad.Q) THEN
    IF fbTrigUp.Q AND (NOT fbTrigDown.Q) THEN
        IF nCvInt < DL_COUNT_MAX THEN
            nCvInt   := nCvInt + 1;
            bUpPulse := TRUE;
        END_IF
    ELSIF fbTrigDown.Q AND (NOT fbTrigUp.Q) THEN
        IF nCvInt > DL_COUNT_MIN THEN
            nCvInt   := nCvInt - 1;
            bDnPulse := TRUE;
        END_IF
    ELSIF fbTrigUp.Q AND fbTrigDown.Q THEN
        IF nCvInt < DL_COUNT_MAX THEN
            nCvInt   := nCvInt + 1;  // 加优先：同拍双边沿净加 1
            bUpPulse := TRUE;
        END_IF
    END_IF
END_IF

(*------------------------------------------------------------------------------
 * 段 8｜饱和标志每拍重算：饱和位不是事件位，而是状态的派生量
 *      Saturation flags recomputed every cycle as derived state
 *-----------------------------------------------------------------------------*)
IF nCvInt >= DL_COUNT_MAX THEN
    bAtMax := TRUE;
ELSE
    bAtMax := FALSE;
END_IF

IF nCvInt <= DL_COUNT_MIN THEN
    bAtMin := TRUE;
ELSE
    bAtMin := FALSE;
END_IF

(*------------------------------------------------------------------------------
 * 段 9｜比较输出每拍重写（R27 保持语义）：禁止只在跨预设那一拍赋值
 *      Comparison outputs rewritten every cycle to keep the holding semantics
 *-----------------------------------------------------------------------------*)
IF bEnable AND (nCvInt >= nPresetUp) THEN
    bQu := TRUE;
ELSE
    bQu := FALSE;
END_IF

IF bEnable AND (nCvInt <= nPresetDn) THEN
    bQd := TRUE;
ELSE
    bQd := FALSE;
END_IF

(*------------------------------------------------------------------------------
 * 段 10｜对外镜像输出：内部值单一来源，外部只读
 *      Mirror the internal count to the output pin, single source of truth
 *-----------------------------------------------------------------------------*)
nCv := nCvInt;

(*------------------------------------------------------------------------------
 * 防御式默认码说明（0216）：本块为计数型，无 CASE 主状态机，故 0216 不参与
 * 正常运行路径，仅作为后续维护者新增分支时的保留码，禁止挪作他用。
 *-----------------------------------------------------------------------------*)
END_FUNCTION_BLOCK

(* ---- FB_DL_MonthWindowCheck.st ---- *)
(*==============================================================================
 * 组件名称 (Component)  : FB_DL_MonthWindowCheck
 * 所属子库 (Sublibrary) : DL_Base
 * 当前版本 (Version)    : 1.0.0
 * 分类     (Category)   : 时间窗判定功能块（Function Block · Date and Timer）
 * 兼容性   (Platform)   : CODESYS 3.5 / TwinCAT 3 / 汇川 InoProShop / Machine Expert
 *                         仅依赖 Standard.library（R_TRIG / MOD / CASE），零厂商方言
 * 功能简介 (Function)   : 月内第 N 天 / 月末倒数第 N 天的日期窗判定（支持窗口
 *                         宽度天数：目标日起连续 n 天）。可选年度模式（仅指定
 *                         月份生效，用于年度保养窗 / 年度盘点窗）。闰年与月长
 *                         规则独立实现（思想与已入库 FC_DL_DayOfWeekCalc 同源，
 *                         本块仅做月长计算、不做星期推导，注释声明同源不调用）；
 *                         日期全部由引脚注入（沿用 R5「时间由引脚注入」修正，
 *                         不读平台时钟，纯组合窗判定 + 开窗边沿脉冲）。
 *                         与已入库 FB_DL_TimeWindowCheck（日内时窗）职责分离：
 *                         本块是日粒度月窗，二者正交不互调。
 * 开源溯源 (Origin)     : 原创实现（参考 LGF 库 Date and Timer 日期时间分类的
 *                         功能域与参数域，来源标签 lgf-datetime），格里高利
 *                         历闰年规则为公开历法定义，仅借分类/参数域/命名，
 *                         clean-room 实现，未复制任何厂商私有库源码。
 * 日期     (Date)       : 2026-11-15 ｜ 作者 (Author): Daoli Library
 * 依赖     (Depends)    : 无 DL_ 内部调用依赖；Standard.library: R_TRIG
 *
 *------------------------------------------------------------------------------
 * 【引脚契约 / Pin contract】
 *   输入 bEnable       : BOOL — 使能，FALSE 时输出复位（bInWindow FALSE、
 *                               bWindowOpen FALSE、nDaysToTarget -1、码清零）；
 *   输入 nYear         : DINT — 当前年份 [公元年]，如 2026，合法域 >= 1；
 *   输入 nMonth        : DINT — 当前月份 [月]，1~12；
 *   输入 nDay          : DINT — 当前日 [日]，1~当月天数；
 *   输入 nTargetDay    : DINT — 目标日 [日]：正数 = 月内第 N 天（1~31）；
 *                               负数 = 月末倒数第 N 天（-1~-31）；0 = 非法；
 *   输入 nWindowDays   : DINT — 窗口宽度 [日]，1~31，目标日起连续 n 天；
 *   输入 bYearly       : BOOL — TRUE = 年度窗：仅生效月份的月内判定开放；
 *   输入 nYearMonth    : DINT — 年度窗生效月份 [月]，1~12（bYearly = FALSE 忽略）；
 *   输出 bInWindow     : BOOL — 当前日在窗口内（保持型，逐拍重算）；
 *   输出 bWindowOpen   : BOOL — 窗口开启单拍脉冲（R25 三律，R_TRIG 无条件刷新）；
 *   输出 nDaysToTarget : DINT — 相对目标日的天数偏移 [日]，窗口内 = 当前日 −
 *                               目标日（首日 0，逐日递增），窗口外固定 -1；
 *   输出 uErrorId      : UDINT — 故障码，0 = 无故障。
 *
 * 【nDaysToTarget 口径声明 / Countdown semantics（判据写死防误解）】
 *   窗口内：nDaysToTarget := nDay − nTargetAbs（窗口首日 = 0，第 k 日 = k−1），
 *   窗口外（含窗口已过、未到、年度模式非生效月、参数非法、未使能）固定 -1。
 *   口径依据规格「窗口外为 -1，窗内为 0 及以上」两条约束联立推导——
 *   「距目标日剩余天数」按目标日锚点偏移实现，保证 0 值必落在窗口首日，
 *   上层以 nDaysToTarget >= 0 判窗内、以 0 判开窗首日，无二义。
 *
 * 【月长与闰年 / Month length and leap year（独立实现声明）】
 *   闰年：能被 4 整除且不能被 100 整除，或能被 400 整除 → 二月 29 天；
 *   月长：1/3/5/7/8/10/12 月 31 天，4/6/9/11 月 30 天，2 月按闰年 28/29；
 *   本规则与已入库 FC_DL_DayOfWeekCalc 的闰年思想同源（公开格里高利历
 *   定义），本块独立实现、不调用该组件（泳道零互相依赖红线）。
 *
 * 【窗口口径 / Window semantics】
 *   窗口 = [nTargetAbs, nTargetAbs + nWindowDays − 1]，右端超过当月天数时
 *   截断到月末（窗口跨月末不跨月，注释写死；截断属口径而非错误，不置码）。
 *   月末倒数口径：nTargetAbs = 当月天数 − |nTargetDay| + 1（倒数第 1 天 =
 *   月末日），|nTargetDay| 超过当月天数时钳位到当月天数（31 在 2 月自动
 *   收缩到 28/29），钳位置信息级码。
 *
 * 【边界防错清单 / Boundary guard list】
 *   B1 nYear < 1 / nMonth 越界（非 1~12）/ nDay 越界（非 1~当月长）/
 *      nTargetDay = 0 → 置 16#0001_0203，bInWindow FALSE，不判定不误报；
 *   B2 nTargetDay 绝对值钳位 1~当月天数（正超钳到月末、负超钳到月长，
 *      钳位先于取负运算，杜绝 DINT 极值取负回绕穿透）；
 *   B3 nWindowDays 钳位 1~31，nYearMonth 钳位 1~12，均置信息级 16#0001_0109；
 *   B4 bYearly = TRUE 且非生效月 → 直接 FALSE 且不置任何故障码（规格写死）；
 *   B5 bWindowOpen 单拍脉冲遵循 R25 三律：R_TRIG 主周期无条件刷新、
 *      边沿基准 bInWindow 单一来源、脉冲仅开窗拍置位下一拍自清；
 *   B6 全部故障码为信息级瞬时型，每拍重算（预清零 + 逐段置位），无锁存。
 *
 * 【单拍标志 R25 三律落地 / One-shot pulse lifecycle】
 *   置位律：bWindowOpen 仅在 bInWindow 由 FALSE 变 TRUE 的扫描拍为 TRUE；
 *   自清律：bInWindow 每拍预清 FALSE 后重算，R_TRIG.Q 无沿自动回落 FALSE；
 *   基准律：边沿基准唯一来源为输出 bInWindow 本身（保持型逐拍重算），
 *   不存在第二份镜像状态，杜绝基准漂移。
 *
 * 【调用示例 / Call example】
 *   「月末倒数第 3 天起开 5 天年度保养窗（仅 12 月生效）」
 *   fbMonthWin(bEnable := TRUE, nYear := 2026, nMonth := 12, nDay := nToday,
 *              nTargetDay := -3, nWindowDays := 5, bYearly := TRUE,
 *              nYearMonth := 12, bInWindow => bMaintWin,
 *              bWindowOpen => bMaintWinOpen, nDaysToTarget => nToTarget,
 *              uErrorId => uWinErr);
 *
 * 【平台移植注意 / Porting notes】
 *   DINT 的 MOD 与负数取负均为 IEC 61131-3 标准语义；本块通过边界 B2 的
 *   「钳位先于取负」次序，保证取负运算的绝对值不超过 31，远离 DINT 极值，
 *   不触发任何平台相关的极值回绕方言。
 *
 * 【工程背景与应用场景 / Background and use cases】
 *   ① 设备月度保养窗：每月 25 日起开 5 天保养允许窗，窗内放行保养工单；
 *   ② 月末盘点窗：月末倒数第 2 天起开 3 天盘点冻结窗，窗内禁止库存异动；
 *   ③ 年度大保养：bYearly = TRUE 且 nYearMonth = 7，仅每年 7 月的指定日段
 *      放行年度检修流程，其余月份自动关闭不报错；
 *   ④ 计量器具月检提醒：nDaysToTarget 从窗口首日 0 起递增，驱动 HMI 上
 *      "窗口第 N 天"提示与窗口末日前的催办逻辑。
 *
 * 【参数组合矩阵 / Parameter combination matrix】
 *   nTargetDay > 0  ：月内第 N 天开窗（正向锚点，1 = 1 日）；
 *   nTargetDay < 0  ：月末倒数第 N 天开窗（反向锚点，-1 = 月末日）；
 *   nWindowDays = 1 ：单日窗（仅目标日当天）；
 *   nWindowDays > 1 ：连续多日窗，右端自动截断到月末；
 *   bYearly = FALSE ：每月都按同参数判定（月度模式）；
 *   bYearly = TRUE  ：仅 nYearMonth 指定月判定，其余月输出全 FALSE 零码。
 *
 * 【典型时序推演 / Typical timing walkthrough】
 *   设 2026-12，nTargetDay = -3，nWindowDays = 5：
 *     目标日 = 31 − 3 + 1 = 29；窗口 = [29, 33] → 截断 [29, 31]；
 *     nDay = 28 → FALSE / -1        （窗前一日）
 *     nDay = 29 → TRUE  / 开窗脉冲 / 0（窗口首日）
 *     nDay = 30 → TRUE  / 无脉冲   / 1
 *     nDay = 31 → TRUE  / 无脉冲   / 2（窗口末日）
 *     nDay = 1（次月）→ FALSE / -1（不跨月，下月按新月长重判）
 *   开窗脉冲仅 29 日当天一拍，次日起 bInWindow 保持 TRUE 而脉冲回落。
 *
 * 【同族职责分离 / Family separation】
 *   FB_DL_TimeWindowCheck：日内时分秒粒度时窗（TOD 比较）；本块：日粒度
 *   月窗（月长/闰年/月内日号），粒度与口径正交；FC_DL_DayOfWeekCalc：
 *   星期推导（思想同源，本块不调用）；三者零互相调用。
 *
 * 红线自检 (Redline)    : R1 零全局变量表/外部变量引用 ✓ ｜ R2 零物理 IO 地址 ✓
 *                         R3 纯 IEC 61131-3 标准运算 ✓ ｜ R4 日期三重校验+钳位
 *                           先于取负+窗口不跨月截断 ✓
 *                         R5 全变量中英双语同行注释 ✓ ｜ R6 月长 CASE 含 ELSE
 *                           兜底；无主状态机（纯组合窗判定，规格豁免）✓
 *                         R7 R_TRIG 主周期无条件刷新（不置于 IF/CASE 内）✓
 *                         R8 月长/月数/窗宽界限全常量化 ✓
 * 验收推演 (Acceptance) :
 *   W1 2026-12，nTargetDay = -3（月末倒数第 3 = 29 日），nWindowDays = 5，
 *      nDay = 29 → bInWindow TRUE，bWindowOpen 单拍 TRUE，nDaysToTarget = 0；
 *   W2 同上 nDay = 31 → bInWindow TRUE（窗口截断到 31），nDaysToTarget = 2；
 *   W3 同上 nDay = 28 → bInWindow FALSE（28 < 29），nDaysToTarget = -1；
 *   W4 2026-02（平年 28 天），nTargetDay = -1 → 目标日 28；nDay = 28 →
 *      bInWindow TRUE，nDaysToTarget = 0；
 *   W5 2028-02（闰年 29 天），nTargetDay = 30 → 钳位 29，置 0109；nDay = 29
 *      → bInWindow TRUE；
 *   W6 bYearly = TRUE，nMonth = 11，nYearMonth = 12 → bInWindow FALSE，
 *      uErrorId = 0（年度过滤不置码）；
 *   W7 nMonth = 13 → 置 0203，bInWindow FALSE；
 *   W8 nTargetDay = 0 → 置 0203，bInWindow FALSE；
 *   W9 bEnable = FALSE → 全输出复位，uErrorId = 0。
 *
 * 【故障码表 / Error code table】
 *   16#0001_0203  日期参数非法：年份 < 1 / 月份非 1~12 / 日非 1~当月长 /
 *                 nTargetDay = 0，本拍不判定，bInWindow FALSE（信息级瞬时码，
 *                 每拍重算；0203 空闲，0201/0202 已被星期/时窗族登记）；
 *   16#0001_0109  参数钳位提示：nTargetDay 绝对值超当月长 / nWindowDays 越界 /
 *                 nYearMonth 越界，按钳位值继续判定（信息级瞬时码，0109 空闲）。
 *
 * 【实现选择 / Implementation choice】
 *   无主状态机：窗判定为纯组合逻辑（参数校验 → 月长解析 → 目标日解析 →
 *   窗口合成 → 区间判定），逐拍全量重算、无跨拍残留状态（除 R_TRIG 内部
 *   边沿基准外），使能撤除即输出复位；月长解析用 CASE nMonth OF 且带 ELSE
 *   兜底（月份虽已在段 2 校验，ELSE 仍拦截非法值，双保险）。
 *
 * 修订历史 (Revision)   :
 *   2026-11-15  v1.0.0  首版落盘（Round 09 · 泳道 A · LGF Date and Timer 组）
 *============================================================================*)
FUNCTION_BLOCK FB_DL_MonthWindowCheck
VAR_INPUT
    bEnable      : BOOL;                   // 使能，FALSE 时输出复位 / Enable, FALSE resets all outputs
    nYear        : DINT;                   // 当前年份 [公元年]，合法域 >= 1 / Current year [calendar year], legal range >= 1
    nMonth       : DINT;                   // 当前月份 [月]，1~12 / Current month [month], 1~12
    nDay         : DINT;                   // 当前日 [日]，1~当月天数 / Current day [day], 1~days in month
    nTargetDay   : DINT;                   // 目标日 [日]，正 = 月内第 N 天，负 = 月末倒数第 N 天，0 非法 / Target day [day], positive = Nth day, negative = Nth day before month end, 0 illegal
    nWindowDays  : DINT := 1;              // 窗口宽度 [日]，1~31，目标日起连续 n 天 / Window width [days], 1~31, consecutive days from target
    bYearly      : BOOL := FALSE;          // TRUE = 年度窗：仅生效月份开放 / TRUE = yearly window, open only in the configured month
    nYearMonth   : DINT := 1;              // 年度窗生效月份 [月]，1~12，非年度模式忽略 / Yearly-window month [month], 1~12, ignored unless yearly
END_VAR
VAR_OUTPUT
    bInWindow    : BOOL;                   // 当前日在窗口内（保持型逐拍重算）/ Today inside the window (held, recomputed each scan)
    bWindowOpen  : BOOL;                   // 窗口开启单拍脉冲（R25 三律）/ Window-open one-shot pulse (R25 three rules)
    nDaysToTarget: DINT := -1;             // 相对目标日天数偏移 [日]，窗内 0 起，窗外 -1 / Day offset relative to target [days], 0+ inside, -1 outside
    uErrorId     : UDINT;                  // 故障码，0 = 无故障 / Error code, 0 = none
END_VAR
VAR
    fbTrigOpen   : R_TRIG;                 // 窗口开启边沿（主周期无条件刷新）/ Window-open edge detector (unconditionally refreshed each scan)
    nMonthLen    : DINT;                   // 当月天数 [日] / Number of days in the current month [days]
    nTargetAbs   : DINT;                   // 目标日绝对日号（月内第 N 天口径）/ Absolute day number of the target (Nth-day-of-month basis)
    nTodayAbs    : DINT;                   // 今日绝对日号（= nDay，口径统一中间量）/ Absolute day number of today (equal to nDay, unified intermediate)
    bValid       : BOOL;                   // 参数合法标志（本拍判定闸门）/ Parameter validity flag (this-scan verdict gate)
    nWinDays     : DINT;                   // 钳位后的窗口宽度 [日] / Clamped window width [days]
    nWinEnd      : DINT;                   // 窗口结束日号（不跨月截断后）/ Window end day number (month-clipped)
    nWinMonth    : DINT;                   // 钳位后的年度窗生效月份 [月] / Clamped yearly-window month [month]
    nBack        : DINT;                   // 月末倒数天数工作副本 [日] / Working copy of days counted back from month end [days]
    bLeap        : BOOL;                   // 闰年标志（当年）/ Leap-year flag of the current year
    nClampMask   : UDINT;                  // 本拍钳位事件累计位图（诊断用）/ Accumulated clamp-event bitmap this scan (for diagnostics)
END_VAR
VAR CONSTANT
    DL_MONTH_MAX : DINT := 12;             // 年度月数上限 [月] / Number of months per year
    DL_DAY_MAX   : DINT := 31;             // 单月最大天数 [日]，窗口宽度上界 / Maximum days per month [days], window width upper bound
    DL_YEAR_MIN  : DINT := 1;              // 合法年份下界 [公元年] / Legal year lower bound [calendar year]
    DL_ERR_DATE  : UDINT := 16#0001_0203;  // 日期参数非法故障码 / Error code for invalid date parameters
    DL_ERR_CLAMP : UDINT := 16#0001_0109;  // 参数钳位提示故障码 / Error code for parameter clamping notice
END_VAR

(*------------------------------------------------------------------------------
 * 段 1｜输出预清零（R25 自清律 + 信息级瞬时码每拍重算）
 *      Output preset clearing (R25 self-clear rule + transient info codes)
 *      全部输出每拍从安全态重建，不残留上拍结果
 *      All outputs rebuilt from safe state each scan, no last-scan residue
 *-----------------------------------------------------------------------------*)
bInWindow    := FALSE;                    // 窗判定预清 FALSE，段 5 合法路径覆盖 / Window verdict preset FALSE, overwritten by stage 5 on legal paths
bWindowOpen  := FALSE;                    // 开窗脉冲预清 FALSE，段 6 边沿覆盖 / Open pulse preset FALSE, overwritten by stage 6 edge
nDaysToTarget:= -1;                       // 天数偏移预置 -1（窗外安全值）/ Day offset preset to -1 (safe outside value)
uErrorId     := 16#0000_0000;             // 故障码预清零，瞬时码逐段置位 / Error code preset to zero, transient codes raised per stage
nClampMask   := 0;                        // 钳位事件位图清零（Clamp bitmap cleared）
bValid       := TRUE;                     // 参数合法性预置通过（Validity preset to pass）
nTodayAbs    := nDay;                     // 今日日号接管输入（Today's day number takes over the input）

(*------------------------------------------------------------------------------
 * 段 2｜参数校验与钳位（边界 B1/B2/B3）
 *      Parameter validation and clamping (guards B1/B2/B3)
 *      校验失败仅置码关闸，不做部分判定，杜绝非法日期误开窗
 *      Failed checks only raise codes and close the gate, never partial verdicts
 *-----------------------------------------------------------------------------*)
IF NOT bEnable THEN
    bValid := FALSE;                       // 未使能：跳过判定，输出保持预清态 / Disabled: skip verdict, outputs stay at preset state
END_IF

IF bValid AND (nYear < DL_YEAR_MIN) THEN
    bValid   := FALSE;                     // 年份非法关闭闸门 / Illegal year closes the gate
    uErrorId := DL_ERR_DATE;               // 置日期参数非法码 / Raise invalid-date code
END_IF

IF bValid AND ((nMonth < 1) OR (nMonth > DL_MONTH_MAX)) THEN
    bValid   := FALSE;                     // 月份非法关闭闸门 / Illegal month closes the gate
    uErrorId := DL_ERR_DATE;               // 置日期参数非法码 / Raise invalid-date code
END_IF

IF bValid AND ((nDay < 1) OR (nDay > DL_DAY_MAX)) THEN
    bValid   := FALSE;                     // 日号粗校验失败（细校验在月长解析后）/ Coarse day check failed (fine check follows month-length parse)
    uErrorId := DL_ERR_DATE;               // 置日期参数非法码 / Raise invalid-date code
END_IF

(*------------------------------------------------------------------------------
 * 段 3｜年度窗生效月钳位（边界 B3/B4）
 *      Yearly-window month clamping (guards B3/B4)
 *   bYearly = FALSE 时 nWinMonth 不使用；bYearly = TRUE 且越界时钳位到 1
 *   并置钳位提示码，保证钳位值本身永远合法，下游无越界分支
 *-----------------------------------------------------------------------------*)
nWinMonth := nYearMonth;                   // 生效月工作副本接管输入 / Working copy takes over the input
IF (nWinMonth < 1) OR (nWinMonth > DL_MONTH_MAX) THEN
    nWinMonth := 1;                        // 钳位到 1 月（Clamp to month 1）
    nClampMask := nClampMask + 1;          // 钳位事件计数（Clamp event counted）
END_IF

(*------------------------------------------------------------------------------
 * 段 4｜月长解析与闰年判定（独立实现，思想与 FC_DL_DayOfWeekCalc 同源）
 *      Month-length parse and leap-year verdict (independent implementation)
 *   闰年：能被 4 整除且非整百年，或能被 400 整除（格里高利历公开定义）
 *   Leap year: divisible by 4 and not by 100, or divisible by 400
 *   CASE nMonth OF 自带 ELSE 兜底：月份已校验，ELSE 属双保险拦截
 *   CASE carries an ELSE fallback: month pre-validated, ELSE is double insurance
 *-----------------------------------------------------------------------------*)
IF bValid THEN
    bLeap := ((nYear MOD 4 = 0) AND (nYear MOD 100 <> 0)) OR (nYear MOD 400 = 0); // 闰年判定 / Leap-year verdict

    CASE nMonth OF                         // 月长查表（Day-length lookup）
    1, 3, 5, 7, 8, 10, 12:                 // 大月 31 天 / Long months with 31 days
        nMonthLen := 31;                   // 31 天（31 days）
    4, 6, 9, 11:                           // 小月 30 天 / Short months with 30 days
        nMonthLen := 30;                   // 30 天（30 days）
    2:                                     // 二月按闰年 28/29 / February by leap year
        IF bLeap THEN
            nMonthLen := 29;               // 闰二月 29 天 / Leap February, 29 days
        ELSE
            nMonthLen := 28;               // 平二月 28 天 / Common February, 28 days
        END_IF
    ELSE                                   // 兜底：非法月份拦截（双保险）/ Fallback: illegal month intercepted (double insurance)
        nMonthLen := 0;                    // 月长清零，后续细校验必失败 / Zero length forces the fine check to fail
        bValid   := FALSE;                 // 关闭判定闸门（Close the verdict gate）
        uErrorId := DL_ERR_DATE;           // 置日期参数非法码 / Raise invalid-date code
    END_CASE

    IF bValid AND ((nDay < 1) OR (nDay > nMonthLen)) THEN
        bValid   := FALSE;                 // 日号细校验：超当月长（如 2 月 30 日）/ Fine day check: beyond month length (e.g. Feb 30)
        uErrorId := DL_ERR_DATE;           // 置日期参数非法码 / Raise invalid-date code
    END_IF
END_IF

(*------------------------------------------------------------------------------
 * 段 5｜目标日解析与窗口合成（边界 B2 + 窗口不跨月）
 *      Target-day parse and window assembly (guard B2 + no cross-month)
 *   正目标日：月内第 N 天，超当月长钳到月末（31 在 2 月自动收缩）；
 *   负目标日：月末倒数第 N 天 = 月长 − |N| + 1，|N| 先钳位再取负，
 *   杜绝 DINT 极值取负回绕穿透；窗口右端超月长截断到月末不置码（口径）。
 *-----------------------------------------------------------------------------*)
IF bValid THEN
    IF nTargetDay = 0 THEN
        bValid   := FALSE;                 // 0 既非正也非负序号，判非法 / Zero is neither a forward nor backward index, deemed illegal
        uErrorId := DL_ERR_DATE;           // 置日期参数非法码 / Raise invalid-date code
    ELSIF nTargetDay > 0 THEN
        IF nTargetDay > nMonthLen THEN     // 正向越当月长 / Forward index beyond month length
            nTargetAbs := nMonthLen;    // 钳到月末（Clamp to month end）
            nClampMask := nClampMask + 1; // 钳位事件计数（Clamp event counted）
        ELSE
            nTargetAbs := nTargetDay;   // 月内第 N 天原值生效 / Nth day of month taken as-is
        END_IF
    ELSE
        IF nTargetDay < -nMonthLen THEN    // 负向绝对值超当月长 / Backward magnitude beyond month length
            nBack := nMonthLen;            // 先钳位（不取负，防极值回绕）/ Clamp first (no negation, no extreme-value wrap)
            nClampMask := nClampMask + 1;  // 钳位事件计数（Clamp event counted）
        ELSE
            nBack := -nTargetDay;          // 安全取负（|N| ≤ 31 远离 DINT 极值）/ Safe negation (magnitude at most 31, far from DINT limits)
        END_IF
        nTargetAbs := nMonthLen - nBack + 1; // 月末倒数口径：倒数第 1 = 月末日 / Backward basis: 1st from end = last day
    END_IF
END_IF

IF bValid THEN
    nWinDays := nWindowDays;               // 窗宽工作副本接管输入 / Window-width working copy takes over the input
    IF nWinDays < 1 THEN
        nWinDays := 1;                     // 下钳 1 天（Clamp to 1 day）
        nClampMask := nClampMask + 1;      // 钳位事件计数（Clamp event counted）
    END_IF
    IF nWinDays > DL_DAY_MAX THEN
        nWinDays := DL_DAY_MAX;            // 上钳 31 天（Clamp to 31 days）
        nClampMask := nClampMask + 1;      // 钳位事件计数（Clamp event counted）
    END_IF

    nWinEnd := nTargetAbs + nWinDays - 1;  // 窗口右端合成 / Window right edge assembled
    IF nWinEnd > nMonthLen THEN
        nWinEnd := nMonthLen;              // 截断到月末，窗口不跨月（口径，不置码）/ Clip to month end, window never crosses months (policy, no code)
    END_IF
END_IF

(*------------------------------------------------------------------------------
 * 段 6｜窗判定与年度过滤（边界 B4）
 *      Window verdict and yearly filtering (guard B4)
 *   年度模式非生效月 → 直接 FALSE 且不置任何码（规格写死）；
 *   窗内 nDaysToTarget := 当前日 − 目标日（首日 0），窗外保持 -1。
 *-----------------------------------------------------------------------------*)
IF bValid THEN
    IF bYearly AND (nMonth <> nWinMonth) THEN
        bInWindow := FALSE;                // 年度过滤：非生效月不开窗 / Yearly filter: window closed outside the configured month
        (* uErrorId 保持 0：年度过滤属口径而非故障 / uErrorId stays 0: filtering is policy, not fault *)
    ELSE
        bInWindow := (nTodayAbs >= nTargetAbs) AND (nTodayAbs <= nWinEnd); // 区间闭判定 / Closed-interval verdict
        IF bInWindow THEN
            nDaysToTarget := nTodayAbs - nTargetAbs; // 窗内偏移：首日 0 逐日递增 / Inside offset: 0 on the first day, +1 per day
        END_IF
    END_IF
    IF nClampMask > 0 THEN
        uErrorId := DL_ERR_CLAMP;          // 存在钳位事件 → 置钳位提示码 / Any clamp event raises the clamp notice code
    END_IF
END_IF

(*------------------------------------------------------------------------------
 * 段 7｜开窗单拍脉冲（R25 三律 + R7 无条件刷新红线）
 *      Window-open one-shot pulse (R25 three rules + R7 unconditional refresh)
 *   R_TRIG 调用置于主体顶层，严禁挪入 IF/CASE 分支（周期安全红线）；
 *   边沿基准唯一来源 bInWindow；脉冲仅开窗拍为 TRUE，下一拍自清。
 *-----------------------------------------------------------------------------*)
fbTrigOpen(CLK := bInWindow);              // 无条件周期刷新（Unconditional per-cycle refresh）
bWindowOpen := fbTrigOpen.Q;               // 开窗拍单拍脉冲，无沿自动回落 / One-shot on the opening scan, falls back without an edge

(*------------------------------------------------------------------------------
 * 段 8｜验收推演索引 / Acceptance walkthrough index
 *   W1 12 月 29 日（倒数第 3 开 5 天窗）→ TRUE / 脉冲一拍 / 偏移 0
 *   W2 12 月 31 日 → TRUE / 偏移 2（窗口截断到 31）
 *   W3 12 月 28 日 → FALSE / 偏移 -1
 *   W4 2026-02-28（平年倒数第 1）→ TRUE / 偏移 0
 *   W5 2028-02 目标 30 → 钳 29 置 0109，29 日 → TRUE
 *   W6 年度模式 11 月非生效月 → FALSE / 码 0
 *   W7 13 月 → 0203；W8 目标 0 → 0203；W9 未使能 → 全复位
 *-----------------------------------------------------------------------------*)
END_FUNCTION_BLOCK
